(* IEC 61131-3 sources: 2026_Projet_YGO_ExcavatriceDragage/TOOLS/TEST_AUTO_CI/RESULTS/L_SIMULATION/tests (part 11) *)

TEST 'TC-T418-INT-010 Desactivation source pendant armement'
nx := 5000; ny := 5000; raw1 := 0; raw2 := 0; previousButton := FALSE; buttonEdges := 0;
bench.Enable := TRUE; bench.HwReal.Operator.JoyXRaw_ANA1 := 5000; bench.HwReal.Operator.JoyYRaw_ANA2 := 5000;
ADVANCE_TIME(10000000); bench(RawPosM1 := raw1, RawPosM2 := raw2);
bench.SimJoystickRight_Fwd_MAINT_Active := TRUE;
ADVANCE_TIME(10000000); bench(RawPosM1 := raw1, RawPosM2 := raw2);
ADVANCE_TIME(10000000); bench(RawPosM1 := raw1, RawPosM2 := raw2);
ADVANCE_TIME(10000000); bench(RawPosM1 := raw1, RawPosM2 := raw2);
ADVANCE_TIME(10000000); bench(RawPosM1 := raw1, RawPosM2 := raw2);
ADVANCE_TIME(10000000); bench(RawPosM1 := raw1, RawPosM2 := raw2);
ASSERT_TRUE(bench.Operator.JoyBtnRaw, 'Armement en cours');
bench.OperatorSourceActive := FALSE;
ADVANCE_TIME(10000000); bench(RawPosM1 := raw1, RawPosM2 := raw2);
ADVANCE_TIME(10000000); bench(RawPosM1 := raw1, RawPosM2 := raw2);
ADVANCE_TIME(10000000); bench(RawPosM1 := raw1, RawPosM2 := raw2);
ADVANCE_TIME(10000000); bench(RawPosM1 := raw1, RawPosM2 := raw2);
ADVANCE_TIME(10000000); bench(RawPosM1 := raw1, RawPosM2 := raw2);
ADVANCE_TIME(10000000); bench(RawPosM1 := raw1, RawPosM2 := raw2);
ADVANCE_TIME(10000000); bench(RawPosM1 := raw1, RawPosM2 := raw2);
ADVANCE_TIME(10000000); bench(RawPosM1 := raw1, RawPosM2 := raw2);
ADVANCE_TIME(10000000); bench(RawPosM1 := raw1, RawPosM2 := raw2);
ADVANCE_TIME(10000000); bench(RawPosM1 := raw1, RawPosM2 := raw2);
ASSERT_FALSE(bench.Operator.JoyBtnRaw, 'Source reelle sans bouton'); ASSERT_EQ(bench.Operator.JoyXRaw_ANA1, 5000, 'Neutre reel');
bench.OperatorSourceActive := TRUE;
ADVANCE_TIME(10000000); bench(RawPosM1 := raw1, RawPosM2 := raw2);
ADVANCE_TIME(10000000); bench(RawPosM1 := raw1, RawPosM2 := raw2);
ADVANCE_TIME(10000000); bench(RawPosM1 := raw1, RawPosM2 := raw2);
ADVANCE_TIME(10000000); bench(RawPosM1 := raw1, RawPosM2 := raw2);
ADVANCE_TIME(10000000); bench(RawPosM1 := raw1, RawPosM2 := raw2);
ADVANCE_TIME(10000000); bench(RawPosM1 := raw1, RawPosM2 := raw2);
ADVANCE_TIME(10000000); bench(RawPosM1 := raw1, RawPosM2 := raw2);
ADVANCE_TIME(10000000); bench(RawPosM1 := raw1, RawPosM2 := raw2);
ADVANCE_TIME(10000000); bench(RawPosM1 := raw1, RawPosM2 := raw2);
ADVANCE_TIME(10000000); bench(RawPosM1 := raw1, RawPosM2 := raw2);
ADVANCE_TIME(10000000); bench(RawPosM1 := raw1, RawPosM2 := raw2);
ADVANCE_TIME(10000000); bench(RawPosM1 := raw1, RawPosM2 := raw2);
ADVANCE_TIME(10000000); bench(RawPosM1 := raw1, RawPosM2 := raw2);
ADVANCE_TIME(10000000); bench(RawPosM1 := raw1, RawPosM2 := raw2);
ADVANCE_TIME(10000000); bench(RawPosM1 := raw1, RawPosM2 := raw2);
ADVANCE_TIME(10000000); bench(RawPosM1 := raw1, RawPosM2 := raw2);
ADVANCE_TIME(10000000); bench(RawPosM1 := raw1, RawPosM2 := raw2);
ADVANCE_TIME(10000000); bench(RawPosM1 := raw1, RawPosM2 := raw2);
ADVANCE_TIME(10000000); bench(RawPosM1 := raw1, RawPosM2 := raw2);
ADVANCE_TIME(10000000); bench(RawPosM1 := raw1, RawPosM2 := raw2);
ADVANCE_TIME(10000000); bench(RawPosM1 := raw1, RawPosM2 := raw2);
ADVANCE_TIME(10000000); bench(RawPosM1 := raw1, RawPosM2 := raw2);
ADVANCE_TIME(10000000); bench(RawPosM1 := raw1, RawPosM2 := raw2);
ADVANCE_TIME(10000000); bench(RawPosM1 := raw1, RawPosM2 := raw2);
ADVANCE_TIME(10000000); bench(RawPosM1 := raw1, RawPosM2 := raw2);
ADVANCE_TIME(10000000); bench(RawPosM1 := raw1, RawPosM2 := raw2);
ADVANCE_TIME(10000000); bench(RawPosM1 := raw1, RawPosM2 := raw2);
ADVANCE_TIME(10000000); bench(RawPosM1 := raw1, RawPosM2 := raw2);
ADVANCE_TIME(10000000); bench(RawPosM1 := raw1, RawPosM2 := raw2);
ADVANCE_TIME(10000000); bench(RawPosM1 := raw1, RawPosM2 := raw2);
ADVANCE_TIME(10000000); bench(RawPosM1 := raw1, RawPosM2 := raw2);
ADVANCE_TIME(10000000); bench(RawPosM1 := raw1, RawPosM2 := raw2);
ADVANCE_TIME(10000000); bench(RawPosM1 := raw1, RawPosM2 := raw2);
ADVANCE_TIME(10000000); bench(RawPosM1 := raw1, RawPosM2 := raw2);
ADVANCE_TIME(10000000); bench(RawPosM1 := raw1, RawPosM2 := raw2);
ADVANCE_TIME(10000000); bench(RawPosM1 := raw1, RawPosM2 := raw2);
ADVANCE_TIME(10000000); bench(RawPosM1 := raw1, RawPosM2 := raw2);
ADVANCE_TIME(10000000); bench(RawPosM1 := raw1, RawPosM2 := raw2);
ADVANCE_TIME(10000000); bench(RawPosM1 := raw1, RawPosM2 := raw2);
ADVANCE_TIME(10000000); bench(RawPosM1 := raw1, RawPosM2 := raw2);
ADVANCE_TIME(10000000); bench(RawPosM1 := raw1, RawPosM2 := raw2);
ADVANCE_TIME(10000000); bench(RawPosM1 := raw1, RawPosM2 := raw2);
ADVANCE_TIME(10000000); bench(RawPosM1 := raw1, RawPosM2 := raw2);
ADVANCE_TIME(10000000); bench(RawPosM1 := raw1, RawPosM2 := raw2);
ADVANCE_TIME(10000000); bench(RawPosM1 := raw1, RawPosM2 := raw2);
ADVANCE_TIME(10000000); bench(RawPosM1 := raw1, RawPosM2 := raw2);
ADVANCE_TIME(10000000); bench(RawPosM1 := raw1, RawPosM2 := raw2);
ADVANCE_TIME(10000000); bench(RawPosM1 := raw1, RawPosM2 := raw2);
ADVANCE_TIME(10000000); bench(RawPosM1 := raw1, RawPosM2 := raw2);
ADVANCE_TIME(10000000); bench(RawPosM1 := raw1, RawPosM2 := raw2);
ADVANCE_TIME(10000000); bench(RawPosM1 := raw1, RawPosM2 := raw2);
ADVANCE_TIME(10000000); bench(RawPosM1 := raw1, RawPosM2 := raw2);
ADVANCE_TIME(10000000); bench(RawPosM1 := raw1, RawPosM2 := raw2);
ADVANCE_TIME(10000000); bench(RawPosM1 := raw1, RawPosM2 := raw2);
ADVANCE_TIME(10000000); bench(RawPosM1 := raw1, RawPosM2 := raw2);
ADVANCE_TIME(10000000); bench(RawPosM1 := raw1, RawPosM2 := raw2);
ADVANCE_TIME(10000000); bench(RawPosM1 := raw1, RawPosM2 := raw2);
ADVANCE_TIME(10000000); bench(RawPosM1 := raw1, RawPosM2 := raw2);
ADVANCE_TIME(10000000); bench(RawPosM1 := raw1, RawPosM2 := raw2);
ADVANCE_TIME(10000000); bench(RawPosM1 := raw1, RawPosM2 := raw2);
ASSERT_FALSE(bench.Operator.JoyBtnRaw, 'Aucun rearmement apres retour de source'); ASSERT_EQ(bench.Operator.JoyXRaw_ANA1, 5000, 'IHM tenue ignoree');
bench.SimJoystickRight_Fwd_MAINT_Active := FALSE;
ADVANCE_TIME(10000000); bench(RawPosM1 := raw1, RawPosM2 := raw2);
bench.SimJoystickRight_Fwd_MAINT_Active := TRUE;
ADVANCE_TIME(10000000); bench(RawPosM1 := raw1, RawPosM2 := raw2);
ASSERT_TRUE(bench.Operator.JoyBtnRaw, 'Nouvel appui apres relachement disponible');
END_TEST

TEST 'TC-T418-INT-011 Desactivation source pendant retour'
nx := 5000; ny := 5000; raw1 := 0; raw2 := 0; previousButton := FALSE; buttonEdges := 0;
bench.Enable := TRUE; bench.HwReal.Operator.JoyXRaw_ANA1 := 5000; bench.HwReal.Operator.JoyYRaw_ANA2 := 5000;
ADVANCE_TIME(10000000); bench(RawPosM1 := raw1, RawPosM2 := raw2);
bench.SimJoystickRight_Fwd_MAINT_Active := TRUE;
ADVANCE_TIME(10000000); bench(RawPosM1 := raw1, RawPosM2 := raw2);
ADVANCE_TIME(10000000); bench(RawPosM1 := raw1, RawPosM2 := raw2);
ADVANCE_TIME(10000000); bench(RawPosM1 := raw1, RawPosM2 := raw2);
ADVANCE_TIME(10000000); bench(RawPosM1 := raw1, RawPosM2 := raw2);
ADVANCE_TIME(10000000); bench(RawPosM1 := raw1, RawPosM2 := raw2);
ADVANCE_TIME(10000000); bench(RawPosM1 := raw1, RawPosM2 := raw2);
ADVANCE_TIME(10000000); bench(RawPosM1 := raw1, RawPosM2 := raw2);
ADVANCE_TIME(10000000); bench(RawPosM1 := raw1, RawPosM2 := raw2);
ADVANCE_TIME(10000000); bench(RawPosM1 := raw1, RawPosM2 := raw2);
ADVANCE_TIME(10000000); bench(RawPosM1 := raw1, RawPosM2 := raw2);
ADVANCE_TIME(10000000); bench(RawPosM1 := raw1, RawPosM2 := raw2);
ADVANCE_TIME(10000000); bench(RawPosM1 := raw1, RawPosM2 := raw2);
ADVANCE_TIME(10000000); bench(RawPosM1 := raw1, RawPosM2 := raw2);
ADVANCE_TIME(10000000); bench(RawPosM1 := raw1, RawPosM2 := raw2);
ADVANCE_TIME(10000000); bench(RawPosM1 := raw1, RawPosM2 := raw2);
ADVANCE_TIME(10000000); bench(RawPosM1 := raw1, RawPosM2 := raw2);
ADVANCE_TIME(10000000); bench(RawPosM1 := raw1, RawPosM2 := raw2);
ADVANCE_TIME(10000000); bench(RawPosM1 := raw1, RawPosM2 := raw2);
ADVANCE_TIME(10000000); bench(RawPosM1 := raw1, RawPosM2 := raw2);
ADVANCE_TIME(10000000); bench(RawPosM1 := raw1, RawPosM2 := raw2);
ADVANCE_TIME(10000000); bench(RawPosM1 := raw1, RawPosM2 := raw2);
ADVANCE_TIME(10000000); bench(RawPosM1 := raw1, RawPosM2 := raw2);
ADVANCE_TIME(10000000); bench(RawPosM1 := raw1, RawPosM2 := raw2);
ADVANCE_TIME(10000000); bench(RawPosM1 := raw1, RawPosM2 := raw2);
ADVANCE_TIME(10000000); bench(RawPosM1 := raw1, RawPosM2 := raw2);
ADVANCE_TIME(10000000); bench(RawPosM1 := raw1, RawPosM2 := raw2);
ADVANCE_TIME(10000000); bench(RawPosM1 := raw1, RawPosM2 := raw2);
ADVANCE_TIME(10000000); bench(RawPosM1 := raw1, RawPosM2 := raw2);
ADVANCE_TIME(10000000); bench(RawPosM1 := raw1, RawPosM2 := raw2);
ADVANCE_TIME(10000000); bench(RawPosM1 := raw1, RawPosM2 := raw2);
ADVANCE_TIME(10000000); bench(RawPosM1 := raw1, RawPosM2 := raw2);
ADVANCE_TIME(10000000); bench(RawPosM1 := raw1, RawPosM2 := raw2);
ADVANCE_TIME(10000000); bench(RawPosM1 := raw1, RawPosM2 := raw2);
ADVANCE_TIME(10000000); bench(RawPosM1 := raw1, RawPosM2 := raw2);
ADVANCE_TIME(10000000); bench(RawPosM1 := raw1, RawPosM2 := raw2);
ADVANCE_TIME(10000000); bench(RawPosM1 := raw1, RawPosM2 := raw2);
ADVANCE_TIME(10000000); bench(RawPosM1 := raw1, RawPosM2 := raw2);
ADVANCE_TIME(10000000); bench(RawPosM1 := raw1, RawPosM2 := raw2);
ADVANCE_TIME(10000000); bench(RawPosM1 := raw1, RawPosM2 := raw2);
ADVANCE_TIME(10000000); bench(RawPosM1 := raw1, RawPosM2 := raw2);
ADVANCE_TIME(10000000); bench(RawPosM1 := raw1, RawPosM2 := raw2);
ADVANCE_TIME(10000000); bench(RawPosM1 := raw1, RawPosM2 := raw2);
ADVANCE_TIME(10000000); bench(RawPosM1 := raw1, RawPosM2 := raw2);
ADVANCE_TIME(10000000); bench(RawPosM1 := raw1, RawPosM2 := raw2);
ADVANCE_TIME(10000000); bench(RawPosM1 := raw1, RawPosM2 := raw2);
ADVANCE_TIME(10000000); bench(RawPosM1 := raw1, RawPosM2 := raw2);
ADVANCE_TIME(10000000); bench(RawPosM1 := raw1, RawPosM2 := raw2);
ADVANCE_TIME(10000000); bench(RawPosM1 := raw1, RawPosM2 := raw2);
ADVANCE_TIME(10000000); bench(RawPosM1 := raw1, RawPosM2 := raw2);
ADVANCE_TIME(10000000); bench(RawPosM1 := raw1, RawPosM2 := raw2);
ADVANCE_TIME(10000000); bench(RawPosM1 := raw1, RawPosM2 := raw2);
ADVANCE_TIME(10000000); bench(RawPosM1 := raw1, RawPosM2 := raw2);
ADVANCE_TIME(10000000); bench(RawPosM1 := raw1, RawPosM2 := raw2);
ADVANCE_TIME(10000000); bench(RawPosM1 := raw1, RawPosM2 := raw2);
ADVANCE_TIME(10000000); bench(RawPosM1 := raw1, RawPosM2 := raw2);
ADVANCE_TIME(10000000); bench(RawPosM1 := raw1, RawPosM2 := raw2);
ADVANCE_TIME(10000000); bench(RawPosM1 := raw1, RawPosM2 := raw2);
ADVANCE_TIME(10000000); bench(RawPosM1 := raw1, RawPosM2 := raw2);
ADVANCE_TIME(10000000); bench(RawPosM1 := raw1, RawPosM2 := raw2);
ADVANCE_TIME(10000000); bench(RawPosM1 := raw1, RawPosM2 := raw2);
ADVANCE_TIME(10000000); bench(RawPosM1 := raw1, RawPosM2 := raw2);
ADVANCE_TIME(10000000); bench(RawPosM1 := raw1, RawPosM2 := raw2);
ADVANCE_TIME(10000000); bench(RawPosM1 := raw1, RawPosM2 := raw2);
ADVANCE_TIME(10000000); bench(RawPosM1 := raw1, RawPosM2 := raw2);
ADVANCE_TIME(10000000); bench(RawPosM1 := raw1, RawPosM2 := raw2);
bench.SimJoystickRight_Fwd_MAINT_Active := FALSE;
ADVANCE_TIME(10000000); bench(RawPosM1 := raw1, RawPosM2 := raw2);
bench.OperatorSourceActive := FALSE;
ADVANCE_TIME(10000000); bench(RawPosM1 := raw1, RawPosM2 := raw2);
bench.SimJoystickLeft_Rev_TREMIE_Active := TRUE; bench.OperatorSourceActive := TRUE;
ADVANCE_TIME(10000000); bench(RawPosM1 := raw1, RawPosM2 := raw2);
ADVANCE_TIME(10000000); bench(RawPosM1 := raw1, RawPosM2 := raw2);
ADVANCE_TIME(10000000); bench(RawPosM1 := raw1, RawPosM2 := raw2);
ADVANCE_TIME(10000000); bench(RawPosM1 := raw1, RawPosM2 := raw2);
ADVANCE_TIME(10000000); bench(RawPosM1 := raw1, RawPosM2 := raw2);
ADVANCE_TIME(10000000); bench(RawPosM1 := raw1, RawPosM2 := raw2);
ADVANCE_TIME(10000000); bench(RawPosM1 := raw1, RawPosM2 := raw2);
ADVANCE_TIME(10000000); bench(RawPosM1 := raw1, RawPosM2 := raw2);
ADVANCE_TIME(10000000); bench(RawPosM1 := raw1, RawPosM2 := raw2);
ADVANCE_TIME(10000000); bench(RawPosM1 := raw1, RawPosM2 := raw2);
ADVANCE_TIME(10000000); bench(RawPosM1 := raw1, RawPosM2 := raw2);
ADVANCE_TIME(10000000); bench(RawPosM1 := raw1, RawPosM2 := raw2);
ADVANCE_TIME(10000000); bench(RawPosM1 := raw1, RawPosM2 := raw2);
ADVANCE_TIME(10000000); bench(RawPosM1 := raw1, RawPosM2 := raw2);
ADVANCE_TIME(10000000); bench(RawPosM1 := raw1, RawPosM2 := raw2);
ADVANCE_TIME(10000000); bench(RawPosM1 := raw1, RawPosM2 := raw2);
ADVANCE_TIME(10000000); bench(RawPosM1 := raw1, RawPosM2 := raw2);
ADVANCE_TIME(10000000); bench(RawPosM1 := raw1, RawPosM2 := raw2);
ADVANCE_TIME(10000000); bench(RawPosM1 := raw1, RawPosM2 := raw2);
ADVANCE_TIME(10000000); bench(RawPosM1 := raw1, RawPosM2 := raw2);
ADVANCE_TIME(10000000); bench(RawPosM1 := raw1, RawPosM2 := raw2);
ADVANCE_TIME(10000000); bench(RawPosM1 := raw1, RawPosM2 := raw2);
ADVANCE_TIME(10000000); bench(RawPosM1 := raw1, RawPosM2 := raw2);
ADVANCE_TIME(10000000); bench(RawPosM1 := raw1, RawPosM2 := raw2);
ADVANCE_TIME(10000000); bench(RawPosM1 := raw1, RawPosM2 := raw2);
ADVANCE_TIME(10000000); bench(RawPosM1 := raw1, RawPosM2 := raw2);
ADVANCE_TIME(10000000); bench(RawPosM1 := raw1, RawPosM2 := raw2);
ADVANCE_TIME(10000000); bench(RawPosM1 := raw1, RawPosM2 := raw2);
ADVANCE_TIME(10000000); bench(RawPosM1 := raw1, RawPosM2 := raw2);
ADVANCE_TIME(10000000); bench(RawPosM1 := raw1, RawPosM2 := raw2);
ADVANCE_TIME(10000000); bench(RawPosM1 := raw1, RawPosM2 := raw2);
ADVANCE_TIME(10000000); bench(RawPosM1 := raw1, RawPosM2 := raw2);
ADVANCE_TIME(10000000); bench(RawPosM1 := raw1, RawPosM2 := raw2);
ADVANCE_TIME(10000000); bench(RawPosM1 := raw1, RawPosM2 := raw2);
ADVANCE_TIME(10000000); bench(RawPosM1 := raw1, RawPosM2 := raw2);
ADVANCE_TIME(10000000); bench(RawPosM1 := raw1, RawPosM2 := raw2);
ADVANCE_TIME(10000000); bench(RawPosM1 := raw1, RawPosM2 := raw2);
ADVANCE_TIME(10000000); bench(RawPosM1 := raw1, RawPosM2 := raw2);
ADVANCE_TIME(10000000); bench(RawPosM1 := raw1, RawPosM2 := raw2);
ADVANCE_TIME(10000000); bench(RawPosM1 := raw1, RawPosM2 := raw2);
ADVANCE_TIME(10000000); bench(RawPosM1 := raw1, RawPosM2 := raw2);
ADVANCE_TIME(10000000); bench(RawPosM1 := raw1, RawPosM2 := raw2);
ADVANCE_TIME(10000000); bench(RawPosM1 := raw1, RawPosM2 := raw2);
ADVANCE_TIME(10000000); bench(RawPosM1 := raw1, RawPosM2 := raw2);
ADVANCE_TIME(10000000); bench(RawPosM1 := raw1, RawPosM2 := raw2);
ADVANCE_TIME(10000000); bench(RawPosM1 := raw1, RawPosM2 := raw2);
ADVANCE_TIME(10000000); bench(RawPosM1 := raw1, RawPosM2 := raw2);
ADVANCE_TIME(10000000); bench(RawPosM1 := raw1, RawPosM2 := raw2);
ADVANCE_TIME(10000000); bench(RawPosM1 := raw1, RawPosM2 := raw2);
ADVANCE_TIME(10000000); bench(RawPosM1 := raw1, RawPosM2 := raw2);
ADVANCE_TIME(10000000); bench(RawPosM1 := raw1, RawPosM2 := raw2);
ADVANCE_TIME(10000000); bench(RawPosM1 := raw1, RawPosM2 := raw2);
ADVANCE_TIME(10000000); bench(RawPosM1 := raw1, RawPosM2 := raw2);
ADVANCE_TIME(10000000); bench(RawPosM1 := raw1, RawPosM2 := raw2);
ADVANCE_TIME(10000000); bench(RawPosM1 := raw1, RawPosM2 := raw2);
ADVANCE_TIME(10000000); bench(RawPosM1 := raw1, RawPosM2 := raw2);
ADVANCE_TIME(10000000); bench(RawPosM1 := raw1, RawPosM2 := raw2);
ADVANCE_TIME(10000000); bench(RawPosM1 := raw1, RawPosM2 := raw2);
ADVANCE_TIME(10000000); bench(RawPosM1 := raw1, RawPosM2 := raw2);
ADVANCE_TIME(10000000); bench(RawPosM1 := raw1, RawPosM2 := raw2);
ASSERT_EQ(bench.Operator.JoyXRaw_ANA1, 5000, 'Retour interrompu ne charge aucun nouveau geste'); ASSERT_FALSE(bench.Operator.JoyBtnRaw, 'Aucun appui differe');
END_TEST

TEST 'TC-T418-INT-012 Source reelle restitue image sans stimuli manuels'
nx := 5000; ny := 5000; raw1 := 0; raw2 := 0; previousButton := FALSE; buttonEdges := 0;
bench.Enable := TRUE; bench.HwReal.Operator.JoyXRaw_ANA1 := 5000; bench.HwReal.Operator.JoyYRaw_ANA2 := 5000;
bench.OperatorSourceActive := FALSE; bench.SimJoystickRawX := 9999; bench.SimJoystickRawY := 1; bench.SimJoystickRawButton := TRUE;
bench.HwReal.Operator.JoyXRaw_ANA1 := 4321; bench.HwReal.Operator.JoyYRaw_ANA2 := 6789; bench.HwReal.Operator.JoyBtnRaw := FALSE; bench.HwReal.Operator.CanBusState := 0;
ADVANCE_TIME(10000000); bench(RawPosM1 := raw1, RawPosM2 := raw2);
ASSERT_EQ(bench.Operator.JoyXRaw_ANA1, 4321, 'X reel exact'); ASSERT_EQ(bench.Operator.JoyYRaw_ANA2, 6789, 'Y reel exact'); ASSERT_FALSE(bench.Operator.JoyBtnRaw, 'Bouton reel exact'); ASSERT_EQ(bench.Operator.CanBusState, 0, 'Diagnostic reel non remplace par RUNNING');
END_TEST

(* ---- test_sim_translation_loop.st ---- *)
(* T417 - rejeu en boucle fermee : FB_Translation REEL (non modifie) + decodeur + FB_Sim_Translation.
   Voir MOCKS/FB_TestLoopTranslation.st (cablage PRG_05 reproduit ; FB_TranslationOutputInterlock et
   FB_Safety_Translation NON reproduits). Un scan = 20 ms simules. Tests de CARACTERISATION : bandes larges,
   gain 0,02 m/(Hz.s) provisoire (T301) ; ce ne sont pas des mesures terrain. *)

TEST 'TC-T417-LOOP-A Rejeu P1 a 20 Hz, demande TENUE apres arrivee : le plafond d approche maintient 20 Hz vers le variateur'
VAR
    loop : FB_TestLoopTranslation;
END_VAR
    loop.HoldRequest := TRUE;
    ADVANCE_TIME(20000000); loop();
    ADVANCE_TIME(20000000); loop();
    ADVANCE_TIME(20000000); loop();
    ADVANCE_TIME(20000000); loop();
    ADVANCE_TIME(20000000); loop();
    ADVANCE_TIME(20000000); loop();
    ADVANCE_TIME(20000000); loop();
    ADVANCE_TIME(20000000); loop();
    ADVANCE_TIME(20000000); loop();
    ADVANCE_TIME(20000000); loop();
    ADVANCE_TIME(20000000); loop();
    ADVANCE_TIME(20000000); loop();
    ADVANCE_TIME(20000000); loop();
    ADVANCE_TIME(20000000); loop();
    ADVANCE_TIME(20000000); loop();
    ADVANCE_TIME(20000000); loop();
    ADVANCE_TIME(20000000); loop();
    ADVANCE_TIME(20000000); loop();
    ADVANCE_TIME(20000000); loop();
    ADVANCE_TIME(20000000); loop();
    ADVANCE_TIME(20000000); loop();
    ADVANCE_TIME(20000000); loop();
    ADVANCE_TIME(20000000); loop();
    ADVANCE_TIME(20000000); loop();
    ADVANCE_TIME(20000000); loop();
    ADVANCE_TIME(20000000); loop();
    ADVANCE_TIME(20000000); loop();
    ADVANCE_TIME(20000000); loop();
    ADVANCE_TIME(20000000); loop();
    ADVANCE_TIME(20000000); loop();
    ADVANCE_TIME(20000000); loop();
    ADVANCE_TIME(20000000); loop();
    ADVANCE_TIME(20000000); loop();
    ADVANCE_TIME(20000000); loop();
    ADVANCE_TIME(20000000); loop();
    ADVANCE_TIME(20000000); loop();
    ADVANCE_TIME(20000000); loop();
    ADVANCE_TIME(20000000); loop();
    ADVANCE_TIME(20000000); loop();
    ADVANCE_TIME(20000000); loop();
    ADVANCE_TIME(20000000); loop();
    ADVANCE_TIME(20000000); loop();
    ADVANCE_TIME(20000000); loop();
    ADVANCE_TIME(20000000); loop();
    ADVANCE_TIME(20000000); loop();
    ADVANCE_TIME(20000000); loop();
    ADVANCE_TIME(20000000); loop();
    ADVANCE_TIME(20000000); loop();
    ADVANCE_TIME(20000000); loop();
    ADVANCE_TIME(20000000); loop();
    ADVANCE_TIME(20000000); loop();
    ADVANCE_TIME(20000000); loop();
    ADVANCE_TIME(20000000); loop();
    ADVANCE_TIME(20000000); loop();
    ADVANCE_TIME(20000000); loop();
    ADVANCE_TIME(20000000); loop();
    ADVANCE_TIME(20000000); loop();
    ADVANCE_TIME(20000000); loop();
    ADVANCE_TIME(20000000); loop();
    ADVANCE_TIME(20000000); loop();
    ADVANCE_TIME(20000000); loop();
    ADVANCE_TIME(20000000); loop();
    ADVANCE_TIME(20000000); loop();
    ADVANCE_TIME(20000000); loop();
    ADVANCE_TIME(20000000); loop();
    ADVANCE_TIME(20000000); loop();
    ADVANCE_TIME(20000000); loop();
    ADVANCE_TIME(20000000); loop();
    ADVANCE_TIME(20000000); loop();
    ADVANCE_TIME(20000000); loop();
    ADVANCE_TIME(20000000); loop();
    ADVANCE_TIME(20000000); loop();
    ADVANCE_TIME(20000000); loop();
    ADVANCE_TIME(20000000); loop();
    ADVANCE_TIME(20000000); loop();
    ADVANCE_TIME(20000000); loop();
    ADVANCE_TIME(20000000); loop();
    ADVANCE_TIME(20000000); loop();
    ADVANCE_TIME(20000000); loop();
    ADVANCE_TIME(20000000); loop();
    ADVANCE_TIME(20000000); loop();
    ADVANCE_TIME(20000000); loop();
    ADVANCE_TIME(20000000); loop();
    ADVANCE_TIME(20000000); loop();
    ADVANCE_TIME(20000000); loop();
    ADVANCE_TIME(20000000); loop();
    ADVANCE_TIME(20000000); loop();
    ADVANCE_TIME(20000000); loop();
    ADVANCE_TIME(20000000); loop();
    ADVANCE_TIME(20000000); loop();
    ADVANCE_TIME(20000000); loop();
    ADVANCE_TIME(20000000); loop();
    ADVANCE_TIME(20000000); loop();
    ADVANCE_TIME(20000000); loop();
    ADVANCE_TIME(20000000); loop();
    ADVANCE_TIME(20000000); loop();
    ADVANCE_TIME(20000000); loop();
    ADVANCE_TIME(20000000); loop();
    ADVANCE_TIME(20000000); loop();
    ADVANCE_TIME(20000000); loop();
    ADVANCE_TIME(20000000); loop();
    ADVANCE_TIME(20000000); loop();
    ADVANCE_TIME(20000000); loop();
    ADVANCE_TIME(20000000); loop();
    ADVANCE_TIME(20000000); loop();
    ADVANCE_TIME(20000000); loop();
    ADVANCE_TIME(20000000); loop();
    ADVANCE_TIME(20000000); loop();
    ADVANCE_TIME(20000000); loop();
    ADVANCE_TIME(20000000); loop();
    ADVANCE_TIME(20000000); loop();
    ADVANCE_TIME(20000000); loop();
    ADVANCE_TIME(20000000); loop();
    ADVANCE_TIME(20000000); loop();
    ADVANCE_TIME(20000000); loop();
    ADVANCE_TIME(20000000); loop();
    ADVANCE_TIME(20000000); loop();
    ADVANCE_TIME(20000000); loop();
    ADVANCE_TIME(20000000); loop();
    ADVANCE_TIME(20000000); loop();
    ADVANCE_TIME(20000000); loop();
    ADVANCE_TIME(20000000); loop();
    ADVANCE_TIME(20000000); loop();
    ADVANCE_TIME(20000000); loop();
    ADVANCE_TIME(20000000); loop();
    ADVANCE_TIME(20000000); loop();
    ADVANCE_TIME(20000000); loop();
    ADVANCE_TIME(20000000); loop();
    ADVANCE_TIME(20000000); loop();
    ADVANCE_TIME(20000000); loop();
    ADVANCE_TIME(20000000); loop();
    ADVANCE_TIME(20000000); loop();
    ADVANCE_TIME(20000000); loop();
    ADVANCE_TIME(20000000); loop();
    ADVANCE_TIME(20000000); loop();
    ADVANCE_TIME(20000000); loop();
    ADVANCE_TIME(20000000); loop();
    ADVANCE_TIME(20000000); loop();
    ADVANCE_TIME(20000000); loop();
    ADVANCE_TIME(20000000); loop();
    ADVANCE_TIME(20000000); loop();
    ADVANCE_TIME(20000000); loop();
    ADVANCE_TIME(20000000); loop();
    ADVANCE_TIME(20000000); loop();
    ADVANCE_TIME(20000000); loop();
    ADVANCE_TIME(20000000); loop();
    ADVANCE_TIME(20000000); loop();
    ADVANCE_TIME(20000000); loop();
    ADVANCE_TIME(20000000); loop();
    ADVANCE_TIME(20000000); loop();
    ADVANCE_TIME(20000000); loop();
    ADVANCE_TIME(20000000); loop();
    ADVANCE_TIME(20000000); loop();
    ADVANCE_TIME(20000000); loop();
    ADVANCE_TIME(20000000); loop();
    ADVANCE_TIME(20000000); loop();
    ADVANCE_TIME(20000000); loop();
    ADVANCE_TIME(20000000); loop();
    ADVANCE_TIME(20000000); loop();
    ADVANCE_TIME(20000000); loop();
    ADVANCE_TIME(20000000); loop();
    ADVANCE_TIME(20000000); loop();
    ADVANCE_TIME(20000000); loop();
    ADVANCE_TIME(20000000); loop();
    ADVANCE_TIME(20000000); loop();
    ADVANCE_TIME(20000000); loop();
    ADVANCE_TIME(20000000); loop();
    ADVANCE_TIME(20000000); loop();
    ADVANCE_TIME(20000000); loop();
    ADVANCE_TIME(20000000); loop();
    ADVANCE_TIME(20000000); loop();
    ADVANCE_TIME(20000000); loop();
    ADVANCE_TIME(20000000); loop();
    ADVANCE_TIME(20000000); loop();
    ADVANCE_TIME(20000000); loop();
    ADVANCE_TIME(20000000); loop();
    ADVANCE_TIME(20000000); loop();
    ADVANCE_TIME(20000000); loop();
    ADVANCE_TIME(20000000); loop();
    ADVANCE_TIME(20000000); loop();
    ADVANCE_TIME(20000000); loop();
    ADVANCE_TIME(20000000); loop();
    ADVANCE_TIME(20000000); loop();
    ADVANCE_TIME(20000000); loop();
    ADVANCE_TIME(20000000); loop();
    ADVANCE_TIME(20000000); loop();
    ADVANCE_TIME(20000000); loop();
    ADVANCE_TIME(20000000); loop();
    ADVANCE_TIME(20000000); loop();
    ADVANCE_TIME(20000000); loop();
    ADVANCE_TIME(20000000); loop();
    ADVANCE_TIME(20000000); loop();
    ADVANCE_TIME(20000000); loop();
    ADVANCE_TIME(20000000); loop();
    ADVANCE_TIME(20000000); loop();
    ADVANCE_TIME(20000000); loop();
    ADVANCE_TIME(20000000); loop();
    ADVANCE_TIME(20000000); loop();
    ADVANCE_TIME(20000000); loop();
    ADVANCE_TIME(20000000); loop();
    ADVANCE_TIME(20000000); loop();
    ADVANCE_TIME(20000000); loop();
    ADVANCE_TIME(20000000); loop();
    ADVANCE_TIME(20000000); loop();
    ADVANCE_TIME(20000000); loop();
    ADVANCE_TIME(20000000); loop();
    ADVANCE_TIME(20000000); loop();
    ADVANCE_TIME(20000000); loop();
    ADVANCE_TIME(20000000); loop();
    ADVANCE_TIME(20000000); loop();
    ADVANCE_TIME(20000000); loop();
    ADVANCE_TIME(20000000); loop();
    ADVANCE_TIME(20000000); loop();
    ADVANCE_TIME(20000000); loop();
    ADVANCE_TIME(20000000); loop();
    ADVANCE_TIME(20000000); loop();
    ADVANCE_TIME(20000000); loop();
    ADVANCE_TIME(20000000); loop();
    ADVANCE_TIME(20000000); loop();
    ADVANCE_TIME(20000000); loop();
    ADVANCE_TIME(20000000); loop();
    ADVANCE_TIME(20000000); loop();
    ADVANCE_TIME(20000000); loop();
    ADVANCE_TIME(20000000); loop();
    ADVANCE_TIME(20000000); loop();
    ADVANCE_TIME(20000000); loop();
    ADVANCE_TIME(20000000); loop();
    ADVANCE_TIME(20000000); loop();
    ADVANCE_TIME(20000000); loop();
    ADVANCE_TIME(20000000); loop();
    ADVANCE_TIME(20000000); loop();
    ADVANCE_TIME(20000000); loop();
    ADVANCE_TIME(20000000); loop();
    ADVANCE_TIME(20000000); loop();
    ADVANCE_TIME(20000000); loop();
    ADVANCE_TIME(20000000); loop();
    ADVANCE_TIME(20000000); loop();
    ADVANCE_TIME(20000000); loop();
    ADVANCE_TIME(20000000); loop();
    ADVANCE_TIME(20000000); loop();
    ADVANCE_TIME(20000000); loop();
    ADVANCE_TIME(20000000); loop();
    ADVANCE_TIME(20000000); loop();
    ADVANCE_TIME(20000000); loop();
    ADVANCE_TIME(20000000); loop();
    ADVANCE_TIME(20000000); loop();
    ADVANCE_TIME(20000000); loop();
    ADVANCE_TIME(20000000); loop();
    ADVANCE_TIME(20000000); loop();
    ADVANCE_TIME(20000000); loop();
    ADVANCE_TIME(20000000); loop();
    ADVANCE_TIME(20000000); loop();
    ADVANCE_TIME(20000000); loop();
    ADVANCE_TIME(20000000); loop();
    ADVANCE_TIME(20000000); loop();
    ADVANCE_TIME(20000000); loop();
    ADVANCE_TIME(20000000); loop();
    ADVANCE_TIME(20000000); loop();
    ADVANCE_TIME(20000000); loop();
    ADVANCE_TIME(20000000); loop();
    ADVANCE_TIME(20000000); loop();
    ADVANCE_TIME(20000000); loop();
    ADVANCE_TIME(20000000); loop();
    ADVANCE_TIME(20000000); loop();
    ADVANCE_TIME(20000000); loop();
    ADVANCE_TIME(20000000); loop();
    ADVANCE_TIME(20000000); loop();
    ADVANCE_TIME(20000000); loop();
    ADVANCE_TIME(20000000); loop();
    ADVANCE_TIME(20000000); loop();
    ADVANCE_TIME(20000000); loop();
    ADVANCE_TIME(20000000); loop();
    ADVANCE_TIME(20000000); loop();
    ADVANCE_TIME(20000000); loop();
    ADVANCE_TIME(20000000); loop();
    ADVANCE_TIME(20000000); loop();
    ADVANCE_TIME(20000000); loop();
    ADVANCE_TIME(20000000); loop();
    ADVANCE_TIME(20000000); loop();
    ADVANCE_TIME(20000000); loop();
    ADVANCE_TIME(20000000); loop();
    ADVANCE_TIME(20000000); loop();
    ADVANCE_TIME(20000000); loop();
    ADVANCE_TIME(20000000); loop();
    ADVANCE_TIME(20000000); loop();
    ADVANCE_TIME(20000000); loop();
    ADVANCE_TIME(20000000); loop();
    ADVANCE_TIME(20000000); loop();
    ADVANCE_TIME(20000000); loop();
    ADVANCE_TIME(20000000); loop();
    ADVANCE_TIME(20000000); loop();
    ADVANCE_TIME(20000000); loop();
    ADVANCE_TIME(20000000); loop();
    ADVANCE_TIME(20000000); loop();
    ADVANCE_TIME(20000000); loop();
    ADVANCE_TIME(20000000); loop();
    ADVANCE_TIME(20000000); loop();
    ADVANCE_TIME(20000000); loop();
    ADVANCE_TIME(20000000); loop();
    ADVANCE_TIME(20000000); loop();
    ADVANCE_TIME(20000000); loop();
    ADVANCE_TIME(20000000); loop();
    ADVANCE_TIME(20000000); loop();
    ADVANCE_TIME(20000000); loop();
    ADVANCE_TIME(20000000); loop();
    ADVANCE_TIME(20000000); loop();
    ADVANCE_TIME(20000000); loop();
    ADVANCE_TIME(20000000); loop();
    ADVANCE_TIME(20000000); loop();
    ADVANCE_TIME(20000000); loop();
    ADVANCE_TIME(20000000); loop();
    ADVANCE_TIME(20000000); loop();
    ADVANCE_TIME(20000000); loop();
    ADVANCE_TIME(20000000); loop();
    ADVANCE_TIME(20000000); loop();
    ADVANCE_TIME(20000000); loop();
    ADVANCE_TIME(20000000); loop();
    ADVANCE_TIME(20000000); loop();
    ADVANCE_TIME(20000000); loop();
    ADVANCE_TIME(20000000); loop();
    ADVANCE_TIME(20000000); loop();
    ADVANCE_TIME(20000000); loop();
    ADVANCE_TIME(20000000); loop();
    ADVANCE_TIME(20000000); loop();
    ADVANCE_TIME(20000000); loop();
    ADVANCE_TIME(20000000); loop();
    ADVANCE_TIME(20000000); loop();
    ADVANCE_TIME(20000000); loop();
    ADVANCE_TIME(20000000); loop();
    ADVANCE_TIME(20000000); loop();
    ADVANCE_TIME(20000000); loop();
    ADVANCE_TIME(20000000); loop();
    ADVANCE_TIME(20000000); loop();
    ADVANCE_TIME(20000000); loop();
    ADVANCE_TIME(20000000); loop();
    ADVANCE_TIME(20000000); loop();
    ADVANCE_TIME(20000000); loop();
    ADVANCE_TIME(20000000); loop();
    ADVANCE_TIME(20000000); loop();
    ADVANCE_TIME(20000000); loop();
    ADVANCE_TIME(20000000); loop();
    ADVANCE_TIME(20000000); loop();
    ADVANCE_TIME(20000000); loop();
    ADVANCE_TIME(20000000); loop();
    ADVANCE_TIME(20000000); loop();
    ADVANCE_TIME(20000000); loop();
    ADVANCE_TIME(20000000); loop();
    ADVANCE_TIME(20000000); loop();
    ADVANCE_TIME(20000000); loop();
    ADVANCE_TIME(20000000); loop();
    ADVANCE_TIME(20000000); loop();
    ADVANCE_TIME(20000000); loop();
    ADVANCE_TIME(20000000); loop();
    ADVANCE_TIME(20000000); loop();
    ADVANCE_TIME(20000000); loop();
    ADVANCE_TIME(20000000); loop();
    ADVANCE_TIME(20000000); loop();
    ADVANCE_TIME(20000000); loop();
    ADVANCE_TIME(20000000); loop();
    ADVANCE_TIME(20000000); loop();
    ADVANCE_TIME(20000000); loop();
    ADVANCE_TIME(20000000); loop();
    ADVANCE_TIME(20000000); loop();
    ADVANCE_TIME(20000000); loop();
    ADVANCE_TIME(20000000); loop();
    ADVANCE_TIME(20000000); loop();
    ADVANCE_TIME(20000000); loop();
    ADVANCE_TIME(20000000); loop();
    ADVANCE_TIME(20000000); loop();
    ADVANCE_TIME(20000000); loop();
    ADVANCE_TIME(20000000); loop();
    ADVANCE_TIME(20000000); loop();
    ADVANCE_TIME(20000000); loop();
    ADVANCE_TIME(20000000); loop();
    ADVANCE_TIME(20000000); loop();
    ADVANCE_TIME(20000000); loop();
    ADVANCE_TIME(20000000); loop();
    ADVANCE_TIME(20000000); loop();
    ADVANCE_TIME(20000000); loop();
    ADVANCE_TIME(20000000); loop();
    ADVANCE_TIME(20000000); loop();
    ADVANCE_TIME(20000000); loop();
    ADVANCE_TIME(20000000); loop();
    ADVANCE_TIME(20000000); loop();
    ADVANCE_TIME(20000000); loop();
    ADVANCE_TIME(20000000); loop();
    ADVANCE_TIME(20000000); loop();
    ADVANCE_TIME(20000000); loop();
    ADVANCE_TIME(20000000); loop();
    ADVANCE_TIME(20000000); loop();
    ADVANCE_TIME(20000000); loop();
    ADVANCE_TIME(20000000); loop();
    ADVANCE_TIME(20000000); loop();
    ADVANCE_TIME(20000000); loop();
    ADVANCE_TIME(20000000); loop();
    ADVANCE_TIME(20000000); loop();
    ADVANCE_TIME(20000000); loop();
    ADVANCE_TIME(20000000); loop();
    ADVANCE_TIME(20000000); loop();
    ADVANCE_TIME(20000000); loop();
    ADVANCE_TIME(20000000); loop();
    ADVANCE_TIME(20000000); loop();
    ADVANCE_TIME(20000000); loop();
    ADVANCE_TIME(20000000); loop();
    ADVANCE_TIME(20000000); loop();
    ADVANCE_TIME(20000000); loop();
    ADVANCE_TIME(20000000); loop();
    ADVANCE_TIME(20000000); loop();
    ADVANCE_TIME(20000000); loop();
    ADVANCE_TIME(20000000); loop();
    ADVANCE_TIME(20000000); loop();
    ADVANCE_TIME(20000000); loop();
    ADVANCE_TIME(20000000); loop();
    ADVANCE_TIME(20000000); loop();
    ADVANCE_TIME(20000000); loop();
    ADVANCE_TIME(20000000); loop();
    ADVANCE_TIME(20000000); loop();
    ADVANCE_TIME(20000000); loop();
    ADVANCE_TIME(20000000); loop();
    ADVANCE_TIME(20000000); loop();
    ADVANCE_TIME(20000000); loop();
    ADVANCE_TIME(20000000); loop();
    ADVANCE_TIME(20000000); loop();
    ADVANCE_TIME(20000000); loop();
    ADVANCE_TIME(20000000); loop();
    ADVANCE_TIME(20000000); loop();
    ADVANCE_TIME(20000000); loop();
    ADVANCE_TIME(20000000); loop();
    ADVANCE_TIME(20000000); loop();
    ADVANCE_TIME(20000000); loop();
    ADVANCE_TIME(20000000); loop();
    ADVANCE_TIME(20000000); loop();
    ADVANCE_TIME(20000000); loop();
    ADVANCE_TIME(20000000); loop();
    ADVANCE_TIME(20000000); loop();
    ADVANCE_TIME(20000000); loop();
    ADVANCE_TIME(20000000); loop();
    ADVANCE_TIME(20000000); loop();
    ADVANCE_TIME(20000000); loop();
    ADVANCE_TIME(20000000); loop();
    ADVANCE_TIME(20000000); loop();
    ADVANCE_TIME(20000000); loop();
    ADVANCE_TIME(20000000); loop();
    ADVANCE_TIME(20000000); loop();
    ADVANCE_TIME(20000000); loop();
    ADVANCE_TIME(20000000); loop();
    ADVANCE_TIME(20000000); loop();
    ADVANCE_TIME(20000000); loop();
    ADVANCE_TIME(20000000); loop();
    ADVANCE_TIME(20000000); loop();
    ADVANCE_TIME(20000000); loop();
    ADVANCE_TIME(20000000); loop();
    ADVANCE_TIME(20000000); loop();
    ADVANCE_TIME(20000000); loop();
    ADVANCE_TIME(20000000); loop();
    ADVANCE_TIME(20000000); loop();
    ADVANCE_TIME(20000000); loop();
    ADVANCE_TIME(20000000); loop();
    ADVANCE_TIME(20000000); loop();
    ADVANCE_TIME(20000000); loop();
    ADVANCE_TIME(20000000); loop();
    ADVANCE_TIME(20000000); loop();
    ADVANCE_TIME(20000000); loop();
    ADVANCE_TIME(20000000); loop();
    ADVANCE_TIME(20000000); loop();
    ADVANCE_TIME(20000000); loop();
    ADVANCE_TIME(20000000); loop();
    ADVANCE_TIME(20000000); loop();
    ADVANCE_TIME(20000000); loop();
    ADVANCE_TIME(20000000); loop();
    ADVANCE_TIME(20000000); loop();
    ADVANCE_TIME(20000000); loop();
    ADVANCE_TIME(20000000); loop();
    ADVANCE_TIME(20000000); loop();
    ADVANCE_TIME(20000000); loop();
    ADVANCE_TIME(20000000); loop();
    ADVANCE_TIME(20000000); loop();
    ADVANCE_TIME(20000000); loop();
    ADVANCE_TIME(20000000); loop();
    ADVANCE_TIME(20000000); loop();
    ADVANCE_TIME(20000000); loop();
    ADVANCE_TIME(20000000); loop();
    ADVANCE_TIME(20000000); loop();
    ADVANCE_TIME(20000000); loop();
    ADVANCE_TIME(20000000); loop();
    ADVANCE_TIME(20000000); loop();
    ADVANCE_TIME(20000000); loop();
    ADVANCE_TIME(20000000); loop();
    ADVANCE_TIME(20000000); loop();
    ADVANCE_TIME(20000000); loop();
    ADVANCE_TIME(20000000); loop();
    ADVANCE_TIME(20000000); loop();
    ADVANCE_TIME(20000000); loop();
    ADVANCE_TIME(20000000); loop();
    ADVANCE_TIME(20000000); loop();
    ADVANCE_TIME(20000000); loop();
    ADVANCE_TIME(20000000); loop();
    ADVANCE_TIME(20000000); loop();
    ADVANCE_TIME(20000000); loop();
    ADVANCE_TIME(20000000); loop();
    ADVANCE_TIME(20000000); loop();
    ADVANCE_TIME(20000000); loop();
    ADVANCE_TIME(20000000); loop();
    ADVANCE_TIME(20000000); loop();
    ADVANCE_TIME(20000000); loop();
    ADVANCE_TIME(20000000); loop();
    ADVANCE_TIME(20000000); loop();
    ADVANCE_TIME(20000000); loop();
    ADVANCE_TIME(20000000); loop();
    ADVANCE_TIME(20000000); loop();
    ADVANCE_TIME(20000000); loop();
    ADVANCE_TIME(20000000); loop();
    ADVANCE_TIME(20000000); loop();
    ADVANCE_TIME(20000000); loop();
    ADVANCE_TIME(20000000); loop();
    ADVANCE_TIME(20000000); loop();
    ADVANCE_TIME(20000000); loop();
    ADVANCE_TIME(20000000); loop();
    ADVANCE_TIME(20000000); loop();
    ADVANCE_TIME(20000000); loop();
    ADVANCE_TIME(20000000); loop();
    ADVANCE_TIME(20000000); loop();
    ADVANCE_TIME(20000000); loop();
    ADVANCE_TIME(20000000); loop();
    ADVANCE_TIME(20000000); loop();
    ADVANCE_TIME(20000000); loop();
    ADVANCE_TIME(20000000); loop();
    ADVANCE_TIME(20000000); loop();
    ADVANCE_TIME(20000000); loop();
    ADVANCE_TIME(20000000); loop();
    ADVANCE_TIME(20000000); loop();
    ADVANCE_TIME(20000000); loop();
    ADVANCE_TIME(20000000); loop();
    ADVANCE_TIME(20000000); loop();
    ADVANCE_TIME(20000000); loop();
    ADVANCE_TIME(20000000); loop();
    ADVANCE_TIME(20000000); loop();
    ADVANCE_TIME(20000000); loop();
    ADVANCE_TIME(20000000); loop();
    ADVANCE_TIME(20000000); loop();
    ADVANCE_TIME(20000000); loop();
    ADVANCE_TIME(20000000); loop();
    ADVANCE_TIME(20000000); loop();
    ADVANCE_TIME(20000000); loop();
    ADVANCE_TIME(20000000); loop();
    ADVANCE_TIME(20000000); loop();
    ADVANCE_TIME(20000000); loop();
    ADVANCE_TIME(20000000); loop();
    ADVANCE_TIME(20000000); loop();
    ADVANCE_TIME(20000000); loop();
    ADVANCE_TIME(20000000); loop();
    ADVANCE_TIME(20000000); loop();
    ADVANCE_TIME(20000000); loop();
    ADVANCE_TIME(20000000); loop();
    ADVANCE_TIME(20000000); loop();
    ADVANCE_TIME(20000000); loop();
    ADVANCE_TIME(20000000); loop();
    ADVANCE_TIME(20000000); loop();
    ADVANCE_TIME(20000000); loop();
    ADVANCE_TIME(20000000); loop();
    ADVANCE_TIME(20000000); loop();
    ADVANCE_TIME(20000000); loop();
    ADVANCE_TIME(20000000); loop();
    ADVANCE_TIME(20000000); loop();
    ADVANCE_TIME(20000000); loop();
    ADVANCE_TIME(20000000); loop();
    ADVANCE_TIME(20000000); loop();
    ADVANCE_TIME(20000000); loop();
    ADVANCE_TIME(20000000); loop();
    ADVANCE_TIME(20000000); loop();
    ADVANCE_TIME(20000000); loop();
    ADVANCE_TIME(20000000); loop();
    ADVANCE_TIME(20000000); loop();
    ADVANCE_TIME(20000000); loop();
    ADVANCE_TIME(20000000); loop();
    ADVANCE_TIME(20000000); loop();
    ADVANCE_TIME(20000000); loop();
    ADVANCE_TIME(20000000); loop();
    ADVANCE_TIME(20000000); loop();
    ADVANCE_TIME(20000000); loop();
    ADVANCE_TIME(20000000); loop();
    ADVANCE_TIME(20000000); loop();
    ADVANCE_TIME(20000000); loop();
    ADVANCE_TIME(20000000); loop();
    ADVANCE_TIME(20000000); loop();
    ADVANCE_TIME(20000000); loop();
    ADVANCE_TIME(20000000); loop();
    ADVANCE_TIME(20000000); loop();
    ADVANCE_TIME(20000000); loop();
    ADVANCE_TIME(20000000); loop();
    ADVANCE_TIME(20000000); loop();
    ADVANCE_TIME(20000000); loop();
    ADVANCE_TIME(20000000); loop();
    ADVANCE_TIME(20000000); loop();
    ADVANCE_TIME(20000000); loop();
    ADVANCE_TIME(20000000); loop();
    ADVANCE_TIME(20000000); loop();
    ADVANCE_TIME(20000000); loop();
    ADVANCE_TIME(20000000); loop();
    ADVANCE_TIME(20000000); loop();
    ADVANCE_TIME(20000000); loop();
    ADVANCE_TIME(20000000); loop();
    ADVANCE_TIME(20000000); loop();
    ADVANCE_TIME(20000000); loop();
    ADVANCE_TIME(20000000); loop();
    ADVANCE_TIME(20000000); loop();
    ADVANCE_TIME(20000000); loop();
    ADVANCE_TIME(20000000); loop();
    ADVANCE_TIME(20000000); loop();
    ADVANCE_TIME(20000000); loop();
    ADVANCE_TIME(20000000); loop();
    ADVANCE_TIME(20000000); loop();
    ADVANCE_TIME(20000000); loop();
    ADVANCE_TIME(20000000); loop();
    ADVANCE_TIME(20000000); loop();
    ADVANCE_TIME(20000000); loop();
    ADVANCE_TIME(20000000); loop();
    ADVANCE_TIME(20000000); loop();
    ADVANCE_TIME(20000000); loop();
    ADVANCE_TIME(20000000); loop();
    ADVANCE_TIME(20000000); loop();
    ADVANCE_TIME(20000000); loop();
    ADVANCE_TIME(20000000); loop();
    ADVANCE_TIME(20000000); loop();
    ADVANCE_TIME(20000000); loop();
    ADVANCE_TIME(20000000); loop();
    ADVANCE_TIME(20000000); loop();
    ADVANCE_TIME(20000000); loop();
    ADVANCE_TIME(20000000); loop();
    ADVANCE_TIME(20000000); loop();
    ADVANCE_TIME(20000000); loop();
    ADVANCE_TIME(20000000); loop();
    ADVANCE_TIME(20000000); loop();
    ADVANCE_TIME(20000000); loop();
    ADVANCE_TIME(20000000); loop();
    ADVANCE_TIME(20000000); loop();
    ADVANCE_TIME(20000000); loop();
    ADVANCE_TIME(20000000); loop();
    ADVANCE_TIME(20000000); loop();
    ADVANCE_TIME(20000000); loop();
    ADVANCE_TIME(20000000); loop();
    ADVANCE_TIME(20000000); loop();
    ADVANCE_TIME(20000000); loop();
    ADVANCE_TIME(20000000); loop();
    ADVANCE_TIME(20000000); loop();
    ADVANCE_TIME(20000000); loop();
    ADVANCE_TIME(20000000); loop();
    ADVANCE_TIME(20000000); loop();
    ADVANCE_TIME(20000000); loop();
    ADVANCE_TIME(20000000); loop();
    ADVANCE_TIME(20000000); loop();
    ADVANCE_TIME(20000000); loop();
    ADVANCE_TIME(20000000); loop();
    ADVANCE_TIME(20000000); loop();
    ADVANCE_TIME(20000000); loop();
    ADVANCE_TIME(20000000); loop();
    ADVANCE_TIME(20000000); loop();
    ADVANCE_TIME(20000000); loop();
    ADVANCE_TIME(20000000); loop();
    ADVANCE_TIME(20000000); loop();
    ADVANCE_TIME(20000000); loop();
    ADVANCE_TIME(20000000); loop();
    ADVANCE_TIME(20000000); loop();
    ADVANCE_TIME(20000000); loop();
    ADVANCE_TIME(20000000); loop();
    ADVANCE_TIME(20000000); loop();
    ADVANCE_TIME(20000000); loop();
    ADVANCE_TIME(20000000); loop();
    ADVANCE_TIME(20000000); loop();
    ADVANCE_TIME(20000000); loop();
    ADVANCE_TIME(20000000); loop();
    ADVANCE_TIME(20000000); loop();
    ADVANCE_TIME(20000000); loop();
    ADVANCE_TIME(20000000); loop();
    ADVANCE_TIME(20000000); loop();
    ADVANCE_TIME(20000000); loop();
    ADVANCE_TIME(20000000); loop();
    ADVANCE_TIME(20000000); loop();
    ADVANCE_TIME(20000000); loop();
    ADVANCE_TIME(20000000); loop();
    ADVANCE_TIME(20000000); loop();
    ADVANCE_TIME(20000000); loop();
    ADVANCE_TIME(20000000); loop();
    ADVANCE_TIME(20000000); loop();
    ADVANCE_TIME(20000000); loop();
    ADVANCE_TIME(20000000); loop();
    ADVANCE_TIME(20000000); loop();
    ADVANCE_TIME(20000000); loop();
    ADVANCE_TIME(20000000); loop();
    ADVANCE_TIME(20000000); loop();
    ADVANCE_TIME(20000000); loop();
    ADVANCE_TIME(20000000); loop();
    ADVANCE_TIME(20000000); loop();
    ADVANCE_TIME(20000000); loop();
    ADVANCE_TIME(20000000); loop();
    ADVANCE_TIME(20000000); loop();
    ADVANCE_TIME(20000000); loop();
    ADVANCE_TIME(20000000); loop();
    ADVANCE_TIME(20000000); loop();
    ADVANCE_TIME(20000000); loop();
    ADVANCE_TIME(20000000); loop();
    ADVANCE_TIME(20000000); loop();
    ADVANCE_TIME(20000000); loop();
    ADVANCE_TIME(20000000); loop();
    ADVANCE_TIME(20000000); loop();
    ADVANCE_TIME(20000000); loop();
    ADVANCE_TIME(20000000); loop();
    ADVANCE_TIME(20000000); loop();
    ADVANCE_TIME(20000000); loop();
    ADVANCE_TIME(20000000); loop();
    ADVANCE_TIME(20000000); loop();
    ADVANCE_TIME(20000000); loop();
    ADVANCE_TIME(20000000); loop();
    ADVANCE_TIME(20000000); loop();
    ADVANCE_TIME(20000000); loop();
    ADVANCE_TIME(20000000); loop();
    ADVANCE_TIME(20000000); loop();
    ADVANCE_TIME(20000000); loop();
    ADVANCE_TIME(20000000); loop();
    ADVANCE_TIME(20000000); loop();
    ADVANCE_TIME(20000000); loop();
    ADVANCE_TIME(20000000); loop();
    ADVANCE_TIME(20000000); loop();
    ADVANCE_TIME(20000000); loop();
    ADVANCE_TIME(20000000); loop();
    ADVANCE_TIME(20000000); loop();
    ADVANCE_TIME(20000000); loop();
    ADVANCE_TIME(20000000); loop();
    ADVANCE_TIME(20000000); loop();
    ADVANCE_TIME(20000000); loop();
    ADVANCE_TIME(20000000); loop();
    ADVANCE_TIME(20000000); loop();
    ADVANCE_TIME(20000000); loop();
    ADVANCE_TIME(20000000); loop();
    ADVANCE_TIME(20000000); loop();
    ADVANCE_TIME(20000000); loop();
    ADVANCE_TIME(20000000); loop();
    ADVANCE_TIME(20000000); loop();
    ADVANCE_TIME(20000000); loop();
    ADVANCE_TIME(20000000); loop();
    ADVANCE_TIME(20000000); loop();
    ADVANCE_TIME(20000000); loop();
    ADVANCE_TIME(20000000); loop();
    ADVANCE_TIME(20000000); loop();
    ADVANCE_TIME(20000000); loop();
    ADVANCE_TIME(20000000); loop();
    ADVANCE_TIME(20000000); loop();
    ADVANCE_TIME(20000000); loop();
    ADVANCE_TIME(20000000); loop();
    ADVANCE_TIME(20000000); loop();
    ADVANCE_TIME(20000000); loop();
    ADVANCE_TIME(20000000); loop();
    ADVANCE_TIME(20000000); loop();
    ADVANCE_TIME(20000000); loop();
    ADVANCE_TIME(20000000); loop();
    ADVANCE_TIME(20000000); loop();
    ADVANCE_TIME(20000000); loop();
    ADVANCE_TIME(20000000); loop();
    ADVANCE_TIME(20000000); loop();
    ADVANCE_TIME(20000000); loop();
    ADVANCE_TIME(20000000); loop();
    ADVANCE_TIME(20000000); loop();
    ADVANCE_TIME(20000000); loop();
    ADVANCE_TIME(20000000); loop();
    ADVANCE_TIME(20000000); loop();
    ADVANCE_TIME(20000000); loop();
    ADVANCE_TIME(20000000); loop();
    ADVANCE_TIME(20000000); loop();
    ADVANCE_TIME(20000000); loop();
    ADVANCE_TIME(20000000); loop();
    ADVANCE_TIME(20000000); loop();
    ADVANCE_TIME(20000000); loop();
    ADVANCE_TIME(20000000); loop();
    ADVANCE_TIME(20000000); loop();
    ADVANCE_TIME(20000000); loop();
    ADVANCE_TIME(20000000); loop();
    ADVANCE_TIME(20000000); loop();
    ADVANCE_TIME(20000000); loop();
    ADVANCE_TIME(20000000); loop();
    ADVANCE_TIME(20000000); loop();
    ADVANCE_TIME(20000000); loop();
    ADVANCE_TIME(20000000); loop();
    ADVANCE_TIME(20000000); loop();
    ADVANCE_TIME(20000000); loop();
    ADVANCE_TIME(20000000); loop();
    ADVANCE_TIME(20000000); loop();
    ADVANCE_TIME(20000000); loop();
    ADVANCE_TIME(20000000); loop();
    ADVANCE_TIME(20000000); loop();
    ADVANCE_TIME(20000000); loop();
    ADVANCE_TIME(20000000); loop();
    ADVANCE_TIME(20000000); loop();
    ADVANCE_TIME(20000000); loop();
    ADVANCE_TIME(20000000); loop();
    ADVANCE_TIME(20000000); loop();
    ADVANCE_TIME(20000000); loop();
    ADVANCE_TIME(20000000); loop();
    ADVANCE_TIME(20000000); loop();
    ADVANCE_TIME(20000000); loop();
    ADVANCE_TIME(20000000); loop();
    ADVANCE_TIME(20000000); loop();
    ADVANCE_TIME(20000000); loop();
    ADVANCE_TIME(20000000); loop();
    ADVANCE_TIME(20000000); loop();
    ADVANCE_TIME(20000000); loop();
    ADVANCE_TIME(20000000); loop();
    ADVANCE_TIME(20000000); loop();
    ADVANCE_TIME(20000000); loop();
    ADVANCE_TIME(20000000); loop();
    ADVANCE_TIME(20000000); loop();
    ADVANCE_TIME(20000000); loop();
    ADVANCE_TIME(20000000); loop();
    ADVANCE_TIME(20000000); loop();
    ADVANCE_TIME(20000000); loop();
    ADVANCE_TIME(20000000); loop();
    ADVANCE_TIME(20000000); loop();
    ADVANCE_TIME(20000000); loop();
    ADVANCE_TIME(20000000); loop();
    ADVANCE_TIME(20000000); loop();
    ADVANCE_TIME(20000000); loop();
    ADVANCE_TIME(20000000); loop();
    ADVANCE_TIME(20000000); loop();
    ADVANCE_TIME(20000000); loop();
    ADVANCE_TIME(20000000); loop();
    ADVANCE_TIME(20000000); loop();
    ADVANCE_TIME(20000000); loop();
    ADVANCE_TIME(20000000); loop();
    ADVANCE_TIME(20000000); loop();
    ADVANCE_TIME(20000000); loop();
    ADVANCE_TIME(20000000); loop();
    ADVANCE_TIME(20000000); loop();
    ADVANCE_TIME(20000000); loop();
    ADVANCE_TIME(20000000); loop();
    ADVANCE_TIME(20000000); loop();
    ADVANCE_TIME(20000000); loop();
    ADVANCE_TIME(20000000); loop();
    ADVANCE_TIME(20000000); loop();
    ADVANCE_TIME(20000000); loop();
    ADVANCE_TIME(20000000); loop();
    ADVANCE_TIME(20000000); loop();
    ADVANCE_TIME(20000000); loop();
    ADVANCE_TIME(20000000); loop();
    ADVANCE_TIME(20000000); loop();
    ADVANCE_TIME(20000000); loop();
    ADVANCE_TIME(20000000); loop();
    ADVANCE_TIME(20000000); loop();
    ADVANCE_TIME(20000000); loop();
    ADVANCE_TIME(20000000); loop();
    ADVANCE_TIME(20000000); loop();
    ADVANCE_TIME(20000000); loop();
    ADVANCE_TIME(20000000); loop();
    ADVANCE_TIME(20000000); loop();
    ADVANCE_TIME(20000000); loop();
    ADVANCE_TIME(20000000); loop();
    ADVANCE_TIME(20000000); loop();
    ADVANCE_TIME(20000000); loop();
    ADVANCE_TIME(20000000); loop();
    ADVANCE_TIME(20000000); loop();
    ADVANCE_TIME(20000000); loop();
    ADVANCE_TIME(20000000); loop();
    ADVANCE_TIME(20000000); loop();
    ADVANCE_TIME(20000000); loop();
    ADVANCE_TIME(20000000); loop();
    ADVANCE_TIME(20000000); loop();
    ADVANCE_TIME(20000000); loop();
    ADVANCE_TIME(20000000); loop();
    ADVANCE_TIME(20000000); loop();
    ADVANCE_TIME(20000000); loop();
    ADVANCE_TIME(20000000); loop();
    ADVANCE_TIME(20000000); loop();
    ADVANCE_TIME(20000000); loop();
    ADVANCE_TIME(20000000); loop();
    ADVANCE_TIME(20000000); loop();
    ADVANCE_TIME(20000000); loop();
    ADVANCE_TIME(20000000); loop();
    ADVANCE_TIME(20000000); loop();
    ADVANCE_TIME(20000000); loop();
    ADVANCE_TIME(20000000); loop();
    ADVANCE_TIME(20000000); loop();
    ADVANCE_TIME(20000000); loop();
    ADVANCE_TIME(20000000); loop();
    ADVANCE_TIME(20000000); loop();
    ADVANCE_TIME(20000000); loop();
    ADVANCE_TIME(20000000); loop();
    ADVANCE_TIME(20000000); loop();
    ADVANCE_TIME(20000000); loop();
    ADVANCE_TIME(20000000); loop();
    ADVANCE_TIME(20000000); loop();
    ADVANCE_TIME(20000000); loop();
    ADVANCE_TIME(20000000); loop();
    ADVANCE_TIME(20000000); loop();
    ADVANCE_TIME(20000000); loop();
    ADVANCE_TIME(20000000); loop();
    ADVANCE_TIME(20000000); loop();
    ADVANCE_TIME(20000000); loop();
    ADVANCE_TIME(20000000); loop();
    ADVANCE_TIME(20000000); loop();
    ADVANCE_TIME(20000000); loop();
    ADVANCE_TIME(20000000); loop();
    ADVANCE_TIME(20000000); loop();
    ADVANCE_TIME(20000000); loop();
    ADVANCE_TIME(20000000); loop();
    ADVANCE_TIME(20000000); loop();
    ADVANCE_TIME(20000000); loop();
    ADVANCE_TIME(20000000); loop();
    ADVANCE_TIME(20000000); loop();
    ADVANCE_TIME(20000000); loop();
    ADVANCE_TIME(20000000); loop();
    ADVANCE_TIME(20000000); loop();
    ADVANCE_TIME(20000000); loop();
    ADVANCE_TIME(20000000); loop();
    ADVANCE_TIME(20000000); loop();
    ADVANCE_TIME(20000000); loop();
    ADVANCE_TIME(20000000); loop();
    ADVANCE_TIME(20000000); loop();
    ADVANCE_TIME(20000000); loop();
    ADVANCE_TIME(20000000); loop();
    ADVANCE_TIME(20000000); loop();
    ADVANCE_TIME(20000000); loop();
    ADVANCE_TIME(20000000); loop();
    ADVANCE_TIME(20000000); loop();
    ADVANCE_TIME(20000000); loop();
    ADVANCE_TIME(20000000); loop();
    ADVANCE_TIME(20000000); loop();
    ADVANCE_TIME(20000000); loop();
    ADVANCE_TIME(20000000); loop();
    ADVANCE_TIME(20000000); loop();
    ADVANCE_TIME(20000000); loop();
    ADVANCE_TIME(20000000); loop();
    ADVANCE_TIME(20000000); loop();
    ADVANCE_TIME(20000000); loop();
    ADVANCE_TIME(20000000); loop();
    ADVANCE_TIME(20000000); loop();
    ADVANCE_TIME(20000000); loop();
    ADVANCE_TIME(20000000); loop();
    ADVANCE_TIME(20000000); loop();
    ADVANCE_TIME(20000000); loop();
    ADVANCE_TIME(20000000); loop();
    ADVANCE_TIME(20000000); loop();
    ADVANCE_TIME(20000000); loop();
    ADVANCE_TIME(20000000); loop();
    ADVANCE_TIME(20000000); loop();
    ADVANCE_TIME(20000000); loop();
    ADVANCE_TIME(20000000); loop();
    ADVANCE_TIME(20000000); loop();
    ADVANCE_TIME(20000000); loop();
    ADVANCE_TIME(20000000); loop();
    ADVANCE_TIME(20000000); loop();
    ADVANCE_TIME(20000000); loop();
    ADVANCE_TIME(20000000); loop();
    ADVANCE_TIME(20000000); loop();
    ADVANCE_TIME(20000000); loop();
    ADVANCE_TIME(20000000); loop();
    ADVANCE_TIME(20000000); loop();
    ADVANCE_TIME(20000000); loop();
    ADVANCE_TIME(20000000); loop();
    ADVANCE_TIME(20000000); loop();
    ADVANCE_TIME(20000000); loop();
    ADVANCE_TIME(20000000); loop();
    ADVANCE_TIME(20000000); loop();
    ADVANCE_TIME(20000000); loop();
    ADVANCE_TIME(20000000); loop();
    ADVANCE_TIME(20000000); loop();
    ADVANCE_TIME(20000000); loop();
    ADVANCE_TIME(20000000); loop();
    ADVANCE_TIME(20000000); loop();
    ADVANCE_TIME(20000000); loop();
    ADVANCE_TIME(20000000); loop();
    ADVANCE_TIME(20000000); loop();
    ADVANCE_TIME(20000000); loop();
    ADVANCE_TIME(20000000); loop();
    ADVANCE_TIME(20000000); loop();
    ADVANCE_TIME(20000000); loop();
    ADVANCE_TIME(20000000); loop();
    ADVANCE_TIME(20000000); loop();
    ADVANCE_TIME(20000000); loop();
    ADVANCE_TIME(20000000); loop();
    ADVANCE_TIME(20000000); loop();
    ADVANCE_TIME(20000000); loop();
    ADVANCE_TIME(20000000); loop();
    ADVANCE_TIME(20000000); loop();
    ADVANCE_TIME(20000000); loop();
    ADVANCE_TIME(20000000); loop();
    ADVANCE_TIME(20000000); loop();
    ADVANCE_TIME(20000000); loop();
    ADVANCE_TIME(20000000); loop();
    ADVANCE_TIME(20000000); loop();
    ADVANCE_TIME(20000000); loop();
    ADVANCE_TIME(20000000); loop();
    ADVANCE_TIME(20000000); loop();
    ADVANCE_TIME(20000000); loop();
    ADVANCE_TIME(20000000); loop();
    ADVANCE_TIME(20000000); loop();
    ADVANCE_TIME(20000000); loop();
    ADVANCE_TIME(20000000); loop();
    ADVANCE_TIME(20000000); loop();
    ADVANCE_TIME(20000000); loop();
    ADVANCE_TIME(20000000); loop();
    ADVANCE_TIME(20000000); loop();
    ADVANCE_TIME(20000000); loop();
    ADVANCE_TIME(20000000); loop();
    ADVANCE_TIME(20000000); loop();
    ADVANCE_TIME(20000000); loop();
    ADVANCE_TIME(20000000); loop();
    ADVANCE_TIME(20000000); loop();
    ADVANCE_TIME(20000000); loop();
    ADVANCE_TIME(20000000); loop();
    ADVANCE_TIME(20000000); loop();
    ADVANCE_TIME(20000000); loop();
    ADVANCE_TIME(20000000); loop();
    ADVANCE_TIME(20000000); loop();
    ADVANCE_TIME(20000000); loop();
    ADVANCE_TIME(20000000); loop();
    ADVANCE_TIME(20000000); loop();
    ADVANCE_TIME(20000000); loop();
    ADVANCE_TIME(20000000); loop();
    ADVANCE_TIME(20000000); loop();
    ADVANCE_TIME(20000000); loop();
    ADVANCE_TIME(20000000); loop();
    ADVANCE_TIME(20000000); loop();
    ADVANCE_TIME(20000000); loop();
    ADVANCE_TIME(20000000); loop();
    ADVANCE_TIME(20000000); loop();
    ADVANCE_TIME(20000000); loop();
    ADVANCE_TIME(20000000); loop();
    ADVANCE_TIME(20000000); loop();
    ADVANCE_TIME(20000000); loop();
    ADVANCE_TIME(20000000); loop();
    ADVANCE_TIME(20000000); loop();
    ADVANCE_TIME(20000000); loop();
    ADVANCE_TIME(20000000); loop();
    ADVANCE_TIME(20000000); loop();
    ADVANCE_TIME(20000000); loop();
    ADVANCE_TIME(20000000); loop();
    ADVANCE_TIME(20000000); loop();
    ADVANCE_TIME(20000000); loop();
    ADVANCE_TIME(20000000); loop();
    ADVANCE_TIME(20000000); loop();
    ADVANCE_TIME(20000000); loop();
    ADVANCE_TIME(20000000); loop();
    ADVANCE_TIME(20000000); loop();
    ADVANCE_TIME(20000000); loop();
    ADVANCE_TIME(20000000); loop();
    ADVANCE_TIME(20000000); loop();
    ADVANCE_TIME(20000000); loop();
    ADVANCE_TIME(20000000); loop();
    ADVANCE_TIME(20000000); loop();
    ADVANCE_TIME(20000000); loop();
    ADVANCE_TIME(20000000); loop();
    ADVANCE_TIME(20000000); loop();
    ADVANCE_TIME(20000000); loop();
    ADVANCE_TIME(20000000); loop();
    ADVANCE_TIME(20000000); loop();
    ADVANCE_TIME(20000000); loop();
    ADVANCE_TIME(20000000); loop();
    ADVANCE_TIME(20000000); loop();
    ADVANCE_TIME(20000000); loop();
    ADVANCE_TIME(20000000); loop();
    ADVANCE_TIME(20000000); loop();
    ADVANCE_TIME(20000000); loop();
    ADVANCE_TIME(20000000); loop();
    ADVANCE_TIME(20000000); loop();
    ADVANCE_TIME(20000000); loop();
    ADVANCE_TIME(20000000); loop();
    ADVANCE_TIME(20000000); loop();
    ADVANCE_TIME(20000000); loop();
    ADVANCE_TIME(20000000); loop();
    ADVANCE_TIME(20000000); loop();
    ADVANCE_TIME(20000000); loop();
    ADVANCE_TIME(20000000); loop();
    ADVANCE_TIME(20000000); loop();
    ADVANCE_TIME(20000000); loop();
    ADVANCE_TIME(20000000); loop();
    ADVANCE_TIME(20000000); loop();
    ADVANCE_TIME(20000000); loop();
    ADVANCE_TIME(20000000); loop();
    ADVANCE_TIME(20000000); loop();
    ADVANCE_TIME(20000000); loop();
    ADVANCE_TIME(20000000); loop();
    ADVANCE_TIME(20000000); loop();
    ADVANCE_TIME(20000000); loop();
    ADVANCE_TIME(20000000); loop();
    ADVANCE_TIME(20000000); loop();
    ADVANCE_TIME(20000000); loop();
    ADVANCE_TIME(20000000); loop();
    ADVANCE_TIME(20000000); loop();
    ADVANCE_TIME(20000000); loop();
    ADVANCE_TIME(20000000); loop();
    ADVANCE_TIME(20000000); loop();
    ADVANCE_TIME(20000000); loop();
    ADVANCE_TIME(20000000); loop();
    ADVANCE_TIME(20000000); loop();
    ADVANCE_TIME(20000000); loop();
    ADVANCE_TIME(20000000); loop();
    ADVANCE_TIME(20000000); loop();
    ADVANCE_TIME(20000000); loop();
    ADVANCE_TIME(20000000); loop();
    ADVANCE_TIME(20000000); loop();
    ADVANCE_TIME(20000000); loop();
    ADVANCE_TIME(20000000); loop();
    ADVANCE_TIME(20000000); loop();
    ADVANCE_TIME(20000000); loop();
    ADVANCE_TIME(20000000); loop();
    ADVANCE_TIME(20000000); loop();
    ADVANCE_TIME(20000000); loop();
    ADVANCE_TIME(20000000); loop();
    ADVANCE_TIME(20000000); loop();
    ADVANCE_TIME(20000000); loop();
    ADVANCE_TIME(20000000); loop();
    ADVANCE_TIME(20000000); loop();
    ADVANCE_TIME(20000000); loop();
    ADVANCE_TIME(20000000); loop();
    ADVANCE_TIME(20000000); loop();
    ADVANCE_TIME(20000000); loop();
    ADVANCE_TIME(20000000); loop();
    ADVANCE_TIME(20000000); loop();
    ADVANCE_TIME(20000000); loop();
    ADVANCE_TIME(20000000); loop();
    ADVANCE_TIME(20000000); loop();
    ADVANCE_TIME(20000000); loop();
    ADVANCE_TIME(20000000); loop();
    ADVANCE_TIME(20000000); loop();
    ADVANCE_TIME(20000000); loop();
    ADVANCE_TIME(20000000); loop();
    ADVANCE_TIME(20000000); loop();
    ADVANCE_TIME(20000000); loop();
    ADVANCE_TIME(20000000); loop();
    ADVANCE_TIME(20000000); loop();
    ADVANCE_TIME(20000000); loop();
    ADVANCE_TIME(20000000); loop();
    ADVANCE_TIME(20000000); loop();
    ADVANCE_TIME(20000000); loop();
    ADVANCE_TIME(20000000); loop();
    ADVANCE_TIME(20000000); loop();
    ADVANCE_TIME(20000000); loop();
    ADVANCE_TIME(20000000); loop();
    ADVANCE_TIME(20000000); loop();
    ADVANCE_TIME(20000000); loop();
    ADVANCE_TIME(20000000); loop();
    ADVANCE_TIME(20000000); loop();
    ADVANCE_TIME(20000000); loop();
    ADVANCE_TIME(20000000); loop();
    ADVANCE_TIME(20000000); loop();
    ADVANCE_TIME(20000000); loop();
    ADVANCE_TIME(20000000); loop();
    ADVANCE_TIME(20000000); loop();
    ADVANCE_TIME(20000000); loop();
    ADVANCE_TIME(20000000); loop();
    ADVANCE_TIME(20000000); loop();
    ADVANCE_TIME(20000000); loop();
    ADVANCE_TIME(20000000); loop();
    ADVANCE_TIME(20000000); loop();
    ADVANCE_TIME(20000000); loop();
    ADVANCE_TIME(20000000); loop();
    ADVANCE_TIME(20000000); loop();
    ADVANCE_TIME(20000000); loop();
    ADVANCE_TIME(20000000); loop();
    ADVANCE_TIME(20000000); loop();
    ADVANCE_TIME(20000000); loop();
    ADVANCE_TIME(20000000); loop();
    ADVANCE_TIME(20000000); loop();
    ADVANCE_TIME(20000000); loop();
    ADVANCE_TIME(20000000); loop();
    ADVANCE_TIME(20000000); loop();
    ADVANCE_TIME(20000000); loop();
    ADVANCE_TIME(20000000); loop();
    ADVANCE_TIME(20000000); loop();
    ADVANCE_TIME(20000000); loop();
    ADVANCE_TIME(20000000); loop();
    ADVANCE_TIME(20000000); loop();
    ADVANCE_TIME(20000000); loop();
    ADVANCE_TIME(20000000); loop();
    ADVANCE_TIME(20000000); loop();
    ADVANCE_TIME(20000000); loop();
    ADVANCE_TIME(20000000); loop();
    ADVANCE_TIME(20000000); loop();
    ADVANCE_TIME(20000000); loop();
    ADVANCE_TIME(20000000); loop();
    ADVANCE_TIME(20000000); loop();
    ADVANCE_TIME(20000000); loop();
    ADVANCE_TIME(20000000); loop();
    ADVANCE_TIME(20000000); loop();
    ADVANCE_TIME(20000000); loop();
    ADVANCE_TIME(20000000); loop();
    ADVANCE_TIME(20000000); loop();
    ADVANCE_TIME(20000000); loop();
    ADVANCE_TIME(20000000); loop();
    ADVANCE_TIME(20000000); loop();
    ADVANCE_TIME(20000000); loop();
    ADVANCE_TIME(20000000); loop();
    ADVANCE_TIME(20000000); loop();
    ADVANCE_TIME(20000000); loop();
    ADVANCE_TIME(20000000); loop();
    ADVANCE_TIME(20000000); loop();
    ADVANCE_TIME(20000000); loop();
    ADVANCE_TIME(20000000); loop();
    ADVANCE_TIME(20000000); loop();
    ADVANCE_TIME(20000000); loop();
    ADVANCE_TIME(20000000); loop();
    ADVANCE_TIME(20000000); loop();
    ADVANCE_TIME(20000000); loop();
    ADVANCE_TIME(20000000); loop();
    ADVANCE_TIME(20000000); loop();
    ADVANCE_TIME(20000000); loop();
    ADVANCE_TIME(20000000); loop();
    ADVANCE_TIME(20000000); loop();
    ADVANCE_TIME(20000000); loop();
    ADVANCE_TIME(20000000); loop();
    ADVANCE_TIME(20000000); loop();
    ADVANCE_TIME(20000000); loop();
    ADVANCE_TIME(20000000); loop();
    ADVANCE_TIME(20000000); loop();
    ADVANCE_TIME(20000000); loop();
    ADVANCE_TIME(20000000); loop();
    ADVANCE_TIME(20000000); loop();
    ADVANCE_TIME(20000000); loop();
    ADVANCE_TIME(20000000); loop();
    ADVANCE_TIME(20000000); loop();
    ADVANCE_TIME(20000000); loop();
    ADVANCE_TIME(20000000); loop();
    ADVANCE_TIME(20000000); loop();
    ADVANCE_TIME(20000000); loop();
    ADVANCE_TIME(20000000); loop();
    ADVANCE_TIME(20000000); loop();
    ADVANCE_TIME(20000000); loop();
    ADVANCE_TIME(20000000); loop();
    ADVANCE_TIME(20000000); loop();
    ADVANCE_TIME(20000000); loop();
    ADVANCE_TIME(20000000); loop();
    ADVANCE_TIME(20000000); loop();
    ADVANCE_TIME(20000000); loop();
    ADVANCE_TIME(20000000); loop();
    ADVANCE_TIME(20000000); loop();
    ADVANCE_TIME(20000000); loop();
    ADVANCE_TIME(20000000); loop();
    ADVANCE_TIME(20000000); loop();
    ADVANCE_TIME(20000000); loop();
    ADVANCE_TIME(20000000); loop();
    ADVANCE_TIME(20000000); loop();
    ADVANCE_TIME(20000000); loop();
    ADVANCE_TIME(20000000); loop();
    ADVANCE_TIME(20000000); loop();
    ADVANCE_TIME(20000000); loop();
    ADVANCE_TIME(20000000); loop();
    ADVANCE_TIME(20000000); loop();
    ADVANCE_TIME(20000000); loop();
    ADVANCE_TIME(20000000); loop();
    ADVANCE_TIME(20000000); loop();
    ADVANCE_TIME(20000000); loop();
    ADVANCE_TIME(20000000); loop();
    ADVANCE_TIME(20000000); loop();
    ADVANCE_TIME(20000000); loop();
    ADVANCE_TIME(20000000); loop();
    ADVANCE_TIME(20000000); loop();
    ADVANCE_TIME(20000000); loop();
    ADVANCE_TIME(20000000); loop();
    ADVANCE_TIME(20000000); loop();
    ADVANCE_TIME(20000000); loop();
    ADVANCE_TIME(20000000); loop();
    ADVANCE_TIME(20000000); loop();
    ADVANCE_TIME(20000000); loop();
    ADVANCE_TIME(20000000); loop();
    ADVANCE_TIME(20000000); loop();
    ADVANCE_TIME(20000000); loop();
    ADVANCE_TIME(20000000); loop();
    ADVANCE_TIME(20000000); loop();
    ADVANCE_TIME(20000000); loop();
    ADVANCE_TIME(20000000); loop();
    ADVANCE_TIME(20000000); loop();
    ADVANCE_TIME(20000000); loop();
    ADVANCE_TIME(20000000); loop();
    ADVANCE_TIME(20000000); loop();
    ADVANCE_TIME(20000000); loop();
    ADVANCE_TIME(20000000); loop();
    ADVANCE_TIME(20000000); loop();
    ADVANCE_TIME(20000000); loop();
    ADVANCE_TIME(20000000); loop();
    ADVANCE_TIME(20000000); loop();
    ADVANCE_TIME(20000000); loop();
    ADVANCE_TIME(20000000); loop();
    ADVANCE_TIME(20000000); loop();
    ADVANCE_TIME(20000000); loop();
    ADVANCE_TIME(20000000); loop();
    ADVANCE_TIME(20000000); loop();
    ADVANCE_TIME(20000000); loop();
    ADVANCE_TIME(20000000); loop();
    ADVANCE_TIME(20000000); loop();
    ADVANCE_TIME(20000000); loop();
    ADVANCE_TIME(20000000); loop();
    ADVANCE_TIME(20000000); loop();
    ADVANCE_TIME(20000000); loop();
    ADVANCE_TIME(20000000); loop();
    ADVANCE_TIME(20000000); loop();
    ADVANCE_TIME(20000000); loop();
    ADVANCE_TIME(20000000); loop();
    ADVANCE_TIME(20000000); loop();
    ADVANCE_TIME(20000000); loop();
    ADVANCE_TIME(20000000); loop();
    ADVANCE_TIME(20000000); loop();
    ADVANCE_TIME(20000000); loop();
    ADVANCE_TIME(20000000); loop();
    ADVANCE_TIME(20000000); loop();
    ADVANCE_TIME(20000000); loop();
    ADVANCE_TIME(20000000); loop();
    ADVANCE_TIME(20000000); loop();
    ADVANCE_TIME(20000000); loop();
    ADVANCE_TIME(20000000); loop();
    ADVANCE_TIME(20000000); loop();
    ADVANCE_TIME(20000000); loop();
    ADVANCE_TIME(20000000); loop();
    ADVANCE_TIME(20000000); loop();
    ADVANCE_TIME(20000000); loop();
    ADVANCE_TIME(20000000); loop();
    ADVANCE_TIME(20000000); loop();
    ADVANCE_TIME(20000000); loop();
    ADVANCE_TIME(20000000); loop();
    ADVANCE_TIME(20000000); loop();
    ADVANCE_TIME(20000000); loop();
    ADVANCE_TIME(20000000); loop();
    ADVANCE_TIME(20000000); loop();
    ADVANCE_TIME(20000000); loop();
    ADVANCE_TIME(20000000); loop();
    ADVANCE_TIME(20000000); loop();
    ADVANCE_TIME(20000000); loop();
    ADVANCE_TIME(20000000); loop();
    ADVANCE_TIME(20000000); loop();
    ADVANCE_TIME(20000000); loop();
    ADVANCE_TIME(20000000); loop();
    ADVANCE_TIME(20000000); loop();
    ADVANCE_TIME(20000000); loop();
    ADVANCE_TIME(20000000); loop();
    ADVANCE_TIME(20000000); loop();
    ADVANCE_TIME(20000000); loop();
    ADVANCE_TIME(20000000); loop();
    ADVANCE_TIME(20000000); loop();
    ADVANCE_TIME(20000000); loop();
    ADVANCE_TIME(20000000); loop();
    ADVANCE_TIME(20000000); loop();
    ADVANCE_TIME(20000000); loop();
    ADVANCE_TIME(20000000); loop();
    ADVANCE_TIME(20000000); loop();
    ADVANCE_TIME(20000000); loop();
    ADVANCE_TIME(20000000); loop();
    ADVANCE_TIME(20000000); loop();
    ADVANCE_TIME(20000000); loop();
    ADVANCE_TIME(20000000); loop();
    ADVANCE_TIME(20000000); loop();
    ADVANCE_TIME(20000000); loop();
    ADVANCE_TIME(20000000); loop();
    ADVANCE_TIME(20000000); loop();
    ADVANCE_TIME(20000000); loop();
    ADVANCE_TIME(20000000); loop();
    ADVANCE_TIME(20000000); loop();
    ADVANCE_TIME(20000000); loop();
    ADVANCE_TIME(20000000); loop();
    ADVANCE_TIME(20000000); loop();
    ADVANCE_TIME(20000000); loop();
    ADVANCE_TIME(20000000); loop();
    ADVANCE_TIME(20000000); loop();
    ADVANCE_TIME(20000000); loop();
    ADVANCE_TIME(20000000); loop();
    ADVANCE_TIME(20000000); loop();
    ADVANCE_TIME(20000000); loop();
    ADVANCE_TIME(20000000); loop();
    ADVANCE_TIME(20000000); loop();
    ADVANCE_TIME(20000000); loop();
    ADVANCE_TIME(20000000); loop();
    ADVANCE_TIME(20000000); loop();
    ADVANCE_TIME(20000000); loop();
    ADVANCE_TIME(20000000); loop();
    ADVANCE_TIME(20000000); loop();
    ADVANCE_TIME(20000000); loop();
    ADVANCE_TIME(20000000); loop();
    ADVANCE_TIME(20000000); loop();
    ADVANCE_TIME(20000000); loop();
    ADVANCE_TIME(20000000); loop();
    ADVANCE_TIME(20000000); loop();
    ADVANCE_TIME(20000000); loop();
    ADVANCE_TIME(20000000); loop();
    ADVANCE_TIME(20000000); loop();
    ADVANCE_TIME(20000000); loop();
    ADVANCE_TIME(20000000); loop();
    ADVANCE_TIME(20000000); loop();
    ADVANCE_TIME(20000000); loop();
    ADVANCE_TIME(20000000); loop();
    ADVANCE_TIME(20000000); loop();
    ADVANCE_TIME(20000000); loop();
    ADVANCE_TIME(20000000); loop();
    ADVANCE_TIME(20000000); loop();
    ADVANCE_TIME(20000000); loop();
    ADVANCE_TIME(20000000); loop();
    ADVANCE_TIME(20000000); loop();
    ADVANCE_TIME(20000000); loop();
    ADVANCE_TIME(20000000); loop();
    ADVANCE_TIME(20000000); loop();
    ADVANCE_TIME(20000000); loop();
    ADVANCE_TIME(20000000); loop();
    ADVANCE_TIME(20000000); loop();
    ADVANCE_TIME(20000000); loop();
    ADVANCE_TIME(20000000); loop();
    ADVANCE_TIME(20000000); loop();
    ADVANCE_TIME(20000000); loop();
    ADVANCE_TIME(20000000); loop();
    ADVANCE_TIME(20000000); loop();
    ADVANCE_TIME(20000000); loop();
    ADVANCE_TIME(20000000); loop();
    ADVANCE_TIME(20000000); loop();
    ADVANCE_TIME(20000000); loop();
    ADVANCE_TIME(20000000); loop();
    ADVANCE_TIME(20000000); loop();
    ADVANCE_TIME(20000000); loop();
    ADVANCE_TIME(20000000); loop();
    ADVANCE_TIME(20000000); loop();
    ADVANCE_TIME(20000000); loop();
    ADVANCE_TIME(20000000); loop();
    ADVANCE_TIME(20000000); loop();
    ADVANCE_TIME(20000000); loop();
    ADVANCE_TIME(20000000); loop();
    ADVANCE_TIME(20000000); loop();
    ADVANCE_TIME(20000000); loop();
    ADVANCE_TIME(20000000); loop();
    ADVANCE_TIME(20000000); loop();
    ADVANCE_TIME(20000000); loop();
    ADVANCE_TIME(20000000); loop();
    ADVANCE_TIME(20000000); loop();
    ADVANCE_TIME(20000000); loop();
    ADVANCE_TIME(20000000); loop();
    ADVANCE_TIME(20000000); loop();
    ADVANCE_TIME(20000000); loop();
    ADVANCE_TIME(20000000); loop();
    ADVANCE_TIME(20000000); loop();
    ADVANCE_TIME(20000000); loop();
    ADVANCE_TIME(20000000); loop();
    ADVANCE_TIME(20000000); loop();
    ADVANCE_TIME(20000000); loop();
    ADVANCE_TIME(20000000); loop();
    ADVANCE_TIME(20000000); loop();
    ADVANCE_TIME(20000000); loop();
    ADVANCE_TIME(20000000); loop();
    ADVANCE_TIME(20000000); loop();
    ADVANCE_TIME(20000000); loop();
    ADVANCE_TIME(20000000); loop();
    ADVANCE_TIME(20000000); loop();
    ADVANCE_TIME(20000000); loop();
    ADVANCE_TIME(20000000); loop();
    ADVANCE_TIME(20000000); loop();
    ADVANCE_TIME(20000000); loop();
    ADVANCE_TIME(20000000); loop();
    ADVANCE_TIME(20000000); loop();
    ADVANCE_TIME(20000000); loop();
    ADVANCE_TIME(20000000); loop();
    ADVANCE_TIME(20000000); loop();
    ADVANCE_TIME(20000000); loop();
    ADVANCE_TIME(20000000); loop();
    ADVANCE_TIME(20000000); loop();
    ADVANCE_TIME(20000000); loop();
    ADVANCE_TIME(20000000); loop();
    ADVANCE_TIME(20000000); loop();
    ADVANCE_TIME(20000000); loop();
    ADVANCE_TIME(20000000); loop();
    ADVANCE_TIME(20000000); loop();
    ADVANCE_TIME(20000000); loop();
    ADVANCE_TIME(20000000); loop();
    ADVANCE_TIME(20000000); loop();
    ADVANCE_TIME(20000000); loop();
    ADVANCE_TIME(20000000); loop();
    ADVANCE_TIME(20000000); loop();
    ADVANCE_TIME(20000000); loop();
    ADVANCE_TIME(20000000); loop();
    ADVANCE_TIME(20000000); loop();
    ADVANCE_TIME(20000000); loop();
    ADVANCE_TIME(20000000); loop();
    ADVANCE_TIME(20000000); loop();
    ADVANCE_TIME(20000000); loop();
    ADVANCE_TIME(20000000); loop();
    ADVANCE_TIME(20000000); loop();
    ADVANCE_TIME(20000000); loop();
    ADVANCE_TIME(20000000); loop();
    ADVANCE_TIME(20000000); loop();
    ADVANCE_TIME(20000000); loop();
    ADVANCE_TIME(20000000); loop();
    ADVANCE_TIME(20000000); loop();
    ADVANCE_TIME(20000000); loop();
    ADVANCE_TIME(20000000); loop();
    ADVANCE_TIME(20000000); loop();
    ADVANCE_TIME(20000000); loop();
    ADVANCE_TIME(20000000); loop();
    ADVANCE_TIME(20000000); loop();
    ADVANCE_TIME(20000000); loop();
    ADVANCE_TIME(20000000); loop();
    ADVANCE_TIME(20000000); loop();
    ADVANCE_TIME(20000000); loop();
    ADVANCE_TIME(20000000); loop();
    ADVANCE_TIME(20000000); loop();
    ADVANCE_TIME(20000000); loop();
    ADVANCE_TIME(20000000); loop();
    ADVANCE_TIME(20000000); loop();
    ADVANCE_TIME(20000000); loop();
    ADVANCE_TIME(20000000); loop();
    ADVANCE_TIME(20000000); loop();
    ADVANCE_TIME(20000000); loop();
    ADVANCE_TIME(20000000); loop();
    ADVANCE_TIME(20000000); loop();
    ADVANCE_TIME(20000000); loop();
    ADVANCE_TIME(20000000); loop();
    ADVANCE_TIME(20000000); loop();
    ADVANCE_TIME(20000000); loop();
    ADVANCE_TIME(20000000); loop();
    ADVANCE_TIME(20000000); loop();
    ADVANCE_TIME(20000000); loop();
    ADVANCE_TIME(20000000); loop();
    ADVANCE_TIME(20000000); loop();
    ADVANCE_TIME(20000000); loop();
    ADVANCE_TIME(20000000); loop();
    ADVANCE_TIME(20000000); loop();
    ADVANCE_TIME(20000000); loop();
    ADVANCE_TIME(20000000); loop();
    ADVANCE_TIME(20000000); loop();
    ADVANCE_TIME(20000000); loop();
    ADVANCE_TIME(20000000); loop();
    ADVANCE_TIME(20000000); loop();
    ADVANCE_TIME(20000000); loop();
    ADVANCE_TIME(20000000); loop();
    ADVANCE_TIME(20000000); loop();
    ADVANCE_TIME(20000000); loop();
    ADVANCE_TIME(20000000); loop();
    ADVANCE_TIME(20000000); loop();
    ADVANCE_TIME(20000000); loop();
    ADVANCE_TIME(20000000); loop();
    ADVANCE_TIME(20000000); loop();
    ADVANCE_TIME(20000000); loop();
    ADVANCE_TIME(20000000); loop();
    ADVANCE_TIME(20000000); loop();
    ADVANCE_TIME(20000000); loop();
    ADVANCE_TIME(20000000); loop();
    ADVANCE_TIME(20000000); loop();
    ADVANCE_TIME(20000000); loop();
    ADVANCE_TIME(20000000); loop();
    ADVANCE_TIME(20000000); loop();
    ADVANCE_TIME(20000000); loop();
    ADVANCE_TIME(20000000); loop();
    ADVANCE_TIME(20000000); loop();
    ADVANCE_TIME(20000000); loop();
    ADVANCE_TIME(20000000); loop();
    ADVANCE_TIME(20000000); loop();
    ADVANCE_TIME(20000000); loop();
    ADVANCE_TIME(20000000); loop();
    ADVANCE_TIME(20000000); loop();
    ADVANCE_TIME(20000000); loop();
    ADVANCE_TIME(20000000); loop();
    ADVANCE_TIME(20000000); loop();
    ADVANCE_TIME(20000000); loop();
    ADVANCE_TIME(20000000); loop();
    ADVANCE_TIME(20000000); loop();
    ADVANCE_TIME(20000000); loop();
    ADVANCE_TIME(20000000); loop();
    ADVANCE_TIME(20000000); loop();
    ADVANCE_TIME(20000000); loop();
    ADVANCE_TIME(20000000); loop();
    ADVANCE_TIME(20000000); loop();
    ADVANCE_TIME(20000000); loop();
    ADVANCE_TIME(20000000); loop();
    ADVANCE_TIME(20000000); loop();
    ADVANCE_TIME(20000000); loop();
    ADVANCE_TIME(20000000); loop();
    ADVANCE_TIME(20000000); loop();
    ADVANCE_TIME(20000000); loop();
    ADVANCE_TIME(20000000); loop();
    ADVANCE_TIME(20000000); loop();
    ADVANCE_TIME(20000000); loop();
    ADVANCE_TIME(20000000); loop();
    ADVANCE_TIME(20000000); loop();
    ADVANCE_TIME(20000000); loop();
    ADVANCE_TIME(20000000); loop();
    ADVANCE_TIME(20000000); loop();
    ADVANCE_TIME(20000000); loop();
    ADVANCE_TIME(20000000); loop();
    ADVANCE_TIME(20000000); loop();
    ADVANCE_TIME(20000000); loop();
    ADVANCE_TIME(20000000); loop();
    ADVANCE_TIME(20000000); loop();
    ADVANCE_TIME(20000000); loop();
    ADVANCE_TIME(20000000); loop();
    ADVANCE_TIME(20000000); loop();
    ADVANCE_TIME(20000000); loop();
    ADVANCE_TIME(20000000); loop();
    ADVANCE_TIME(20000000); loop();
    ADVANCE_TIME(20000000); loop();
    ADVANCE_TIME(20000000); loop();
    ADVANCE_TIME(20000000); loop();
    ADVANCE_TIME(20000000); loop();
    ADVANCE_TIME(20000000); loop();
    ADVANCE_TIME(20000000); loop();
    ADVANCE_TIME(20000000); loop();
    ADVANCE_TIME(20000000); loop();
    ADVANCE_TIME(20000000); loop();
    ADVANCE_TIME(20000000); loop();
    ADVANCE_TIME(20000000); loop();
    ADVANCE_TIME(20000000); loop();
    ADVANCE_TIME(20000000); loop();
    ADVANCE_TIME(20000000); loop();
    ADVANCE_TIME(20000000); loop();
    ADVANCE_TIME(20000000); loop();
    ADVANCE_TIME(20000000); loop();
    ADVANCE_TIME(20000000); loop();
    ADVANCE_TIME(20000000); loop();
    ADVANCE_TIME(20000000); loop();
    ADVANCE_TIME(20000000); loop();
    ADVANCE_TIME(20000000); loop();
    ADVANCE_TIME(20000000); loop();
    ADVANCE_TIME(20000000); loop();
    ADVANCE_TIME(20000000); loop();
    ADVANCE_TIME(20000000); loop();
    ADVANCE_TIME(20000000); loop();
    ADVANCE_TIME(20000000); loop();
    ADVANCE_TIME(20000000); loop();
    ADVANCE_TIME(20000000); loop();
    ADVANCE_TIME(20000000); loop();
    ADVANCE_TIME(20000000); loop();
    ADVANCE_TIME(20000000); loop();
    ADVANCE_TIME(20000000); loop();
    ADVANCE_TIME(20000000); loop();
    ADVANCE_TIME(20000000); loop();
    ADVANCE_TIME(20000000); loop();
    ADVANCE_TIME(20000000); loop();
    ADVANCE_TIME(20000000); loop();
    ADVANCE_TIME(20000000); loop();
    ADVANCE_TIME(20000000); loop();
    ADVANCE_TIME(20000000); loop();
    ADVANCE_TIME(20000000); loop();
    ADVANCE_TIME(20000000); loop();
    ADVANCE_TIME(20000000); loop();
    ADVANCE_TIME(20000000); loop();
    ADVANCE_TIME(20000000); loop();
    ADVANCE_TIME(20000000); loop();
    ADVANCE_TIME(20000000); loop();
    ADVANCE_TIME(20000000); loop();
    ADVANCE_TIME(20000000); loop();
    ADVANCE_TIME(20000000); loop();
    ADVANCE_TIME(20000000); loop();
    ADVANCE_TIME(20000000); loop();
    ADVANCE_TIME(20000000); loop();
    ADVANCE_TIME(20000000); loop();
    ADVANCE_TIME(20000000); loop();
    ADVANCE_TIME(20000000); loop();
    ADVANCE_TIME(20000000); loop();
    ADVANCE_TIME(20000000); loop();
    ADVANCE_TIME(20000000); loop();
    ADVANCE_TIME(20000000); loop();
    ADVANCE_TIME(20000000); loop();
    ADVANCE_TIME(20000000); loop();
    ADVANCE_TIME(20000000); loop();
    ADVANCE_TIME(20000000); loop();
    ADVANCE_TIME(20000000); loop();
    ADVANCE_TIME(20000000); loop();
    ADVANCE_TIME(20000000); loop();
    ADVANCE_TIME(20000000); loop();
    ADVANCE_TIME(20000000); loop();
    ADVANCE_TIME(20000000); loop();
    ADVANCE_TIME(20000000); loop();
    ADVANCE_TIME(20000000); loop();
    ADVANCE_TIME(20000000); loop();
    ADVANCE_TIME(20000000); loop();
    ADVANCE_TIME(20000000); loop();
    ADVANCE_TIME(20000000); loop();
    ADVANCE_TIME(20000000); loop();
    ADVANCE_TIME(20000000); loop();
    ADVANCE_TIME(20000000); loop();
    ADVANCE_TIME(20000000); loop();
    ADVANCE_TIME(20000000); loop();
    ADVANCE_TIME(20000000); loop();
    ADVANCE_TIME(20000000); loop();
    ADVANCE_TIME(20000000); loop();
    ADVANCE_TIME(20000000); loop();
    ADVANCE_TIME(20000000); loop();
    ADVANCE_TIME(20000000); loop();
    ADVANCE_TIME(20000000); loop();
    ADVANCE_TIME(20000000); loop();
    ADVANCE_TIME(20000000); loop();
    ADVANCE_TIME(20000000); loop();
    ADVANCE_TIME(20000000); loop();
    ADVANCE_TIME(20000000); loop();
    ADVANCE_TIME(20000000); loop();
    ADVANCE_TIME(20000000); loop();
    ADVANCE_TIME(20000000); loop();
    ADVANCE_TIME(20000000); loop();
    ADVANCE_TIME(20000000); loop();
    ADVANCE_TIME(20000000); loop();
    ADVANCE_TIME(20000000); loop();
    ADVANCE_TIME(20000000); loop();
    ADVANCE_TIME(20000000); loop();
    ADVANCE_TIME(20000000); loop();
    ADVANCE_TIME(20000000); loop();
    ADVANCE_TIME(20000000); loop();
    ADVANCE_TIME(20000000); loop();
    ADVANCE_TIME(20000000); loop();
    ADVANCE_TIME(20000000); loop();
    ADVANCE_TIME(20000000); loop();
    ADVANCE_TIME(20000000); loop();
    ADVANCE_TIME(20000000); loop();
    ADVANCE_TIME(20000000); loop();
    ADVANCE_TIME(20000000); loop();
    ADVANCE_TIME(20000000); loop();
    ADVANCE_TIME(20000000); loop();
    ADVANCE_TIME(20000000); loop();
    ADVANCE_TIME(20000000); loop();
    ADVANCE_TIME(20000000); loop();
    ADVANCE_TIME(20000000); loop();
    ADVANCE_TIME(20000000); loop();
    ADVANCE_TIME(20000000); loop();
    ADVANCE_TIME(20000000); loop();
    ADVANCE_TIME(20000000); loop();
    ADVANCE_TIME(20000000); loop();
    ADVANCE_TIME(20000000); loop();
    ADVANCE_TIME(20000000); loop();
    ADVANCE_TIME(20000000); loop();
    ADVANCE_TIME(20000000); loop();
    ADVANCE_TIME(20000000); loop();
    ADVANCE_TIME(20000000); loop();
    ADVANCE_TIME(20000000); loop();
    ADVANCE_TIME(20000000); loop();
    ADVANCE_TIME(20000000); loop();
    ADVANCE_TIME(20000000); loop();
    ADVANCE_TIME(20000000); loop();
    ADVANCE_TIME(20000000); loop();
    ADVANCE_TIME(20000000); loop();
    ADVANCE_TIME(20000000); loop();
    ADVANCE_TIME(20000000); loop();
    ADVANCE_TIME(20000000); loop();
    ADVANCE_TIME(20000000); loop();
    ADVANCE_TIME(20000000); loop();
    ADVANCE_TIME(20000000); loop();
    ADVANCE_TIME(20000000); loop();
    ADVANCE_TIME(20000000); loop();
    ADVANCE_TIME(20000000); loop();
    ADVANCE_TIME(20000000); loop();
    ADVANCE_TIME(20000000); loop();
    ADVANCE_TIME(20000000); loop();
    ADVANCE_TIME(20000000); loop();
    ADVANCE_TIME(20000000); loop();
    ADVANCE_TIME(20000000); loop();
    ADVANCE_TIME(20000000); loop();
    ADVANCE_TIME(20000000); loop();
    ADVANCE_TIME(20000000); loop();
    ADVANCE_TIME(20000000); loop();
    ADVANCE_TIME(20000000); loop();
    ADVANCE_TIME(20000000); loop();
    ADVANCE_TIME(20000000); loop();
    ADVANCE_TIME(20000000); loop();
    ADVANCE_TIME(20000000); loop();
    ADVANCE_TIME(20000000); loop();
    ADVANCE_TIME(20000000); loop();
    ADVANCE_TIME(20000000); loop();
    ADVANCE_TIME(20000000); loop();
    ADVANCE_TIME(20000000); loop();
    ADVANCE_TIME(20000000); loop();
    ADVANCE_TIME(20000000); loop();
    ADVANCE_TIME(20000000); loop();
    ADVANCE_TIME(20000000); loop();
    ADVANCE_TIME(20000000); loop();
    ADVANCE_TIME(20000000); loop();
    ADVANCE_TIME(20000000); loop();
    ADVANCE_TIME(20000000); loop();
    ADVANCE_TIME(20000000); loop();
    ADVANCE_TIME(20000000); loop();
    ADVANCE_TIME(20000000); loop();
    ADVANCE_TIME(20000000); loop();
    ADVANCE_TIME(20000000); loop();
    ADVANCE_TIME(20000000); loop();
    ADVANCE_TIME(20000000); loop();
    ADVANCE_TIME(20000000); loop();
    ADVANCE_TIME(20000000); loop();
    ADVANCE_TIME(20000000); loop();
    ADVANCE_TIME(20000000); loop();
    ADVANCE_TIME(20000000); loop();
    ADVANCE_TIME(20000000); loop();
    ADVANCE_TIME(20000000); loop();
    ADVANCE_TIME(20000000); loop();
    ADVANCE_TIME(20000000); loop();
    ADVANCE_TIME(20000000); loop();
    ADVANCE_TIME(20000000); loop();
    ADVANCE_TIME(20000000); loop();
    ADVANCE_TIME(20000000); loop();
    ADVANCE_TIME(20000000); loop();
    ADVANCE_TIME(20000000); loop();
    ADVANCE_TIME(20000000); loop();
    ADVANCE_TIME(20000000); loop();
    ADVANCE_TIME(20000000); loop();
    ADVANCE_TIME(20000000); loop();
    ADVANCE_TIME(20000000); loop();
    ADVANCE_TIME(20000000); loop();
    ADVANCE_TIME(20000000); loop();
    ADVANCE_TIME(20000000); loop();
    ADVANCE_TIME(20000000); loop();
    ADVANCE_TIME(20000000); loop();
    ADVANCE_TIME(20000000); loop();
    ADVANCE_TIME(20000000); loop();
    ADVANCE_TIME(20000000); loop();
    ADVANCE_TIME(20000000); loop();
    ADVANCE_TIME(20000000); loop();
    ADVANCE_TIME(20000000); loop();
    ADVANCE_TIME(20000000); loop();
    ADVANCE_TIME(20000000); loop();
    ADVANCE_TIME(20000000); loop();
    ADVANCE_TIME(20000000); loop();
    ADVANCE_TIME(20000000); loop();
    ADVANCE_TIME(20000000); loop();
    ADVANCE_TIME(20000000); loop();
    ADVANCE_TIME(20000000); loop();
    ADVANCE_TIME(20000000); loop();
    ADVANCE_TIME(20000000); loop();
    ADVANCE_TIME(20000000); loop();
    ADVANCE_TIME(20000000); loop();
    ADVANCE_TIME(20000000); loop();
    ADVANCE_TIME(20000000); loop();
    ADVANCE_TIME(20000000); loop();
    ADVANCE_TIME(20000000); loop();
    ADVANCE_TIME(20000000); loop();
    ADVANCE_TIME(20000000); loop();
    ADVANCE_TIME(20000000); loop();
    ADVANCE_TIME(20000000); loop();
    ADVANCE_TIME(20000000); loop();
    ADVANCE_TIME(20000000); loop();
    ADVANCE_TIME(20000000); loop();
    ADVANCE_TIME(20000000); loop();
    ADVANCE_TIME(20000000); loop();
    ADVANCE_TIME(20000000); loop();
    ADVANCE_TIME(20000000); loop();
    ADVANCE_TIME(20000000); loop();
    ADVANCE_TIME(20000000); loop();
    ADVANCE_TIME(20000000); loop();
    ADVANCE_TIME(20000000); loop();
    ADVANCE_TIME(20000000); loop();
    ADVANCE_TIME(20000000); loop();
    ADVANCE_TIME(20000000); loop();
    ADVANCE_TIME(20000000); loop();
    ADVANCE_TIME(20000000); loop();
    ADVANCE_TIME(20000000); loop();
    ADVANCE_TIME(20000000); loop();
    ADVANCE_TIME(20000000); loop();
    ADVANCE_TIME(20000000); loop();
    ADVANCE_TIME(20000000); loop();
    ADVANCE_TIME(20000000); loop();
    ADVANCE_TIME(20000000); loop();
    ADVANCE_TIME(20000000); loop();
    ADVANCE_TIME(20000000); loop();
    ADVANCE_TIME(20000000); loop();
    ADVANCE_TIME(20000000); loop();
    ADVANCE_TIME(20000000); loop();
    ADVANCE_TIME(20000000); loop();
    ADVANCE_TIME(20000000); loop();
    ADVANCE_TIME(20000000); loop();
    ADVANCE_TIME(20000000); loop();
    ADVANCE_TIME(20000000); loop();
    ADVANCE_TIME(20000000); loop();
    ADVANCE_TIME(20000000); loop();
    ADVANCE_TIME(20000000); loop();
    ADVANCE_TIME(20000000); loop();
    ADVANCE_TIME(20000000); loop();
    ADVANCE_TIME(20000000); loop();
    ADVANCE_TIME(20000000); loop();
    ADVANCE_TIME(20000000); loop();
    ADVANCE_TIME(20000000); loop();
    ADVANCE_TIME(20000000); loop();
    ADVANCE_TIME(20000000); loop();
    ADVANCE_TIME(20000000); loop();
    ADVANCE_TIME(20000000); loop();
    ADVANCE_TIME(20000000); loop();
    ADVANCE_TIME(20000000); loop();
    ADVANCE_TIME(20000000); loop();
    ADVANCE_TIME(20000000); loop();
    ADVANCE_TIME(20000000); loop();
    ADVANCE_TIME(20000000); loop();
    ADVANCE_TIME(20000000); loop();
    ADVANCE_TIME(20000000); loop();
    ADVANCE_TIME(20000000); loop();
    ADVANCE_TIME(20000000); loop();
    ADVANCE_TIME(20000000); loop();
    ADVANCE_TIME(20000000); loop();
    ADVANCE_TIME(20000000); loop();
    ADVANCE_TIME(20000000); loop();
    ADVANCE_TIME(20000000); loop();
    ADVANCE_TIME(20000000); loop();
    ADVANCE_TIME(20000000); loop();
    ADVANCE_TIME(20000000); loop();
    ADVANCE_TIME(20000000); loop();
    ADVANCE_TIME(20000000); loop();
    ADVANCE_TIME(20000000); loop();
    ADVANCE_TIME(20000000); loop();
    ADVANCE_TIME(20000000); loop();
    ADVANCE_TIME(20000000); loop();
    ADVANCE_TIME(20000000); loop();
    ADVANCE_TIME(20000000); loop();
    ADVANCE_TIME(20000000); loop();
    ADVANCE_TIME(20000000); loop();
    ADVANCE_TIME(20000000); loop();
    ADVANCE_TIME(20000000); loop();
    ADVANCE_TIME(20000000); loop();
    ADVANCE_TIME(20000000); loop();
    ADVANCE_TIME(20000000); loop();
    ADVANCE_TIME(20000000); loop();
    ADVANCE_TIME(20000000); loop();
    ADVANCE_TIME(20000000); loop();
    ADVANCE_TIME(20000000); loop();
    ADVANCE_TIME(20000000); loop();
    ADVANCE_TIME(20000000); loop();
    ADVANCE_TIME(20000000); loop();
    ADVANCE_TIME(20000000); loop();
    ADVANCE_TIME(20000000); loop();
    ADVANCE_TIME(20000000); loop();
    ADVANCE_TIME(20000000); loop();
    ADVANCE_TIME(20000000); loop();
    ADVANCE_TIME(20000000); loop();
    ADVANCE_TIME(20000000); loop();
    ADVANCE_TIME(20000000); loop();
    ADVANCE_TIME(20000000); loop();
    ADVANCE_TIME(20000000); loop();
    ADVANCE_TIME(20000000); loop();
    ADVANCE_TIME(20000000); loop();
    ADVANCE_TIME(20000000); loop();
    ADVANCE_TIME(20000000); loop();
    ADVANCE_TIME(20000000); loop();
    ADVANCE_TIME(20000000); loop();
    ADVANCE_TIME(20000000); loop();
    ADVANCE_TIME(20000000); loop();
    ADVANCE_TIME(20000000); loop();
    ADVANCE_TIME(20000000); loop();
    ADVANCE_TIME(20000000); loop();
    ADVANCE_TIME(20000000); loop();
    ADVANCE_TIME(20000000); loop();
    ADVANCE_TIME(20000000); loop();
    ADVANCE_TIME(20000000); loop();
    ADVANCE_TIME(20000000); loop();
    ADVANCE_TIME(20000000); loop();
    ADVANCE_TIME(20000000); loop();
    ADVANCE_TIME(20000000); loop();
    ADVANCE_TIME(20000000); loop();
    ADVANCE_TIME(20000000); loop();
    ADVANCE_TIME(20000000); loop();
    ADVANCE_TIME(20000000); loop();
    ADVANCE_TIME(20000000); loop();
    ADVANCE_TIME(20000000); loop();
    ADVANCE_TIME(20000000); loop();
    ADVANCE_TIME(20000000); loop();
    ADVANCE_TIME(20000000); loop();
    ADVANCE_TIME(20000000); loop();
    ADVANCE_TIME(20000000); loop();
    ADVANCE_TIME(20000000); loop();
    ADVANCE_TIME(20000000); loop();
    ADVANCE_TIME(20000000); loop();
    ADVANCE_TIME(20000000); loop();
    ADVANCE_TIME(20000000); loop();
    ADVANCE_TIME(20000000); loop();
    ADVANCE_TIME(20000000); loop();
    ADVANCE_TIME(20000000); loop();
    ADVANCE_TIME(20000000); loop();
    ADVANCE_TIME(20000000); loop();
    ADVANCE_TIME(20000000); loop();
    ADVANCE_TIME(20000000); loop();
    ADVANCE_TIME(20000000); loop();
    ADVANCE_TIME(20000000); loop();
    ADVANCE_TIME(20000000); loop();
    ADVANCE_TIME(20000000); loop();
    ADVANCE_TIME(20000000); loop();
    ADVANCE_TIME(20000000); loop();
    ADVANCE_TIME(20000000); loop();
    ADVANCE_TIME(20000000); loop();
    ADVANCE_TIME(20000000); loop();
    ADVANCE_TIME(20000000); loop();
    ADVANCE_TIME(20000000); loop();
    ADVANCE_TIME(20000000); loop();
    ADVANCE_TIME(20000000); loop();
    ADVANCE_TIME(20000000); loop();
    ADVANCE_TIME(20000000); loop();
    ADVANCE_TIME(20000000); loop();
    ADVANCE_TIME(20000000); loop();
    ADVANCE_TIME(20000000); loop();
    ADVANCE_TIME(20000000); loop();
    ADVANCE_TIME(20000000); loop();
    ADVANCE_TIME(20000000); loop();
    ADVANCE_TIME(20000000); loop();
    ADVANCE_TIME(20000000); loop();
    ADVANCE_TIME(20000000); loop();
    ADVANCE_TIME(20000000); loop();
    ADVANCE_TIME(20000000); loop();
    ADVANCE_TIME(20000000); loop();
    ADVANCE_TIME(20000000); loop();
    ADVANCE_TIME(20000000); loop();
    ADVANCE_TIME(20000000); loop();
    ADVANCE_TIME(20000000); loop();
    ADVANCE_TIME(20000000); loop();
    ADVANCE_TIME(20000000); loop();
    ADVANCE_TIME(20000000); loop();
    ADVANCE_TIME(20000000); loop();
    ADVANCE_TIME(20000000); loop();
    ADVANCE_TIME(20000000); loop();
    ADVANCE_TIME(20000000); loop();
    ADVANCE_TIME(20000000); loop();
    ADVANCE_TIME(20000000); loop();
    ADVANCE_TIME(20000000); loop();
    ADVANCE_TIME(20000000); loop();
    ADVANCE_TIME(20000000); loop();
    ADVANCE_TIME(20000000); loop();
    ADVANCE_TIME(20000000); loop();
    ADVANCE_TIME(20000000); loop();
    ADVANCE_TIME(20000000); loop();
    ADVANCE_TIME(20000000); loop();
    ADVANCE_TIME(20000000); loop();
    ADVANCE_TIME(20000000); loop();
    ADVANCE_TIME(20000000); loop();
    ADVANCE_TIME(20000000); loop();
    ADVANCE_TIME(20000000); loop();
    ADVANCE_TIME(20000000); loop();
    ADVANCE_TIME(20000000); loop();
    ADVANCE_TIME(20000000); loop();
    ADVANCE_TIME(20000000); loop();
    ADVANCE_TIME(20000000); loop();
    ADVANCE_TIME(20000000); loop();
    ADVANCE_TIME(20000000); loop();
    ADVANCE_TIME(20000000); loop();
    ADVANCE_TIME(20000000); loop();
    ADVANCE_TIME(20000000); loop();
    ADVANCE_TIME(20000000); loop();
    ADVANCE_TIME(20000000); loop();
    ADVANCE_TIME(20000000); loop();
    ADVANCE_TIME(20000000); loop();
    ADVANCE_TIME(20000000); loop();
    ADVANCE_TIME(20000000); loop();
    ADVANCE_TIME(20000000); loop();
    ADVANCE_TIME(20000000); loop();
    ADVANCE_TIME(20000000); loop();
    ADVANCE_TIME(20000000); loop();
    ADVANCE_TIME(20000000); loop();
    ADVANCE_TIME(20000000); loop();
    ADVANCE_TIME(20000000); loop();
    ADVANCE_TIME(20000000); loop();
    ADVANCE_TIME(20000000); loop();
    ADVANCE_TIME(20000000); loop();
    ADVANCE_TIME(20000000); loop();
    ADVANCE_TIME(20000000); loop();
    ADVANCE_TIME(20000000); loop();
    ADVANCE_TIME(20000000); loop();
    ADVANCE_TIME(20000000); loop();
    ADVANCE_TIME(20000000); loop();
    ADVANCE_TIME(20000000); loop();
    ADVANCE_TIME(20000000); loop();
    ADVANCE_TIME(20000000); loop();
    ADVANCE_TIME(20000000); loop();
    ADVANCE_TIME(20000000); loop();
    ADVANCE_TIME(20000000); loop();
    ADVANCE_TIME(20000000); loop();
    ADVANCE_TIME(20000000); loop();
    ADVANCE_TIME(20000000); loop();
    ADVANCE_TIME(20000000); loop();
    ADVANCE_TIME(20000000); loop();
    ADVANCE_TIME(20000000); loop();
    ADVANCE_TIME(20000000); loop();
    ADVANCE_TIME(20000000); loop();
    ADVANCE_TIME(20000000); loop();
    ADVANCE_TIME(20000000); loop();
    ADVANCE_TIME(20000000); loop();
    ADVANCE_TIME(20000000); loop();
    ADVANCE_TIME(20000000); loop();
    ADVANCE_TIME(20000000); loop();
    ADVANCE_TIME(20000000); loop();
    ADVANCE_TIME(20000000); loop();
    ADVANCE_TIME(20000000); loop();
    ADVANCE_TIME(20000000); loop();
    ADVANCE_TIME(20000000); loop();
    ADVANCE_TIME(20000000); loop();
    ADVANCE_TIME(20000000); loop();
    ADVANCE_TIME(20000000); loop();
    ADVANCE_TIME(20000000); loop();
    ADVANCE_TIME(20000000); loop();
    ADVANCE_TIME(20000000); loop();
    ADVANCE_TIME(20000000); loop();
    ADVANCE_TIME(20000000); loop();
    ADVANCE_TIME(20000000); loop();
    ADVANCE_TIME(20000000); loop();
    ADVANCE_TIME(20000000); loop();
    ADVANCE_TIME(20000000); loop();
    ADVANCE_TIME(20000000); loop();
    ADVANCE_TIME(20000000); loop();
    ADVANCE_TIME(20000000); loop();
    ADVANCE_TIME(20000000); loop();
    ADVANCE_TIME(20000000); loop();
    ADVANCE_TIME(20000000); loop();
    ADVANCE_TIME(20000000); loop();
    ADVANCE_TIME(20000000); loop();
    ADVANCE_TIME(20000000); loop();
    ADVANCE_TIME(20000000); loop();
    ADVANCE_TIME(20000000); loop();
    ADVANCE_TIME(20000000); loop();
    ADVANCE_TIME(20000000); loop();
    ADVANCE_TIME(20000000); loop();
    ADVANCE_TIME(20000000); loop();
    ADVANCE_TIME(20000000); loop();
    ADVANCE_TIME(20000000); loop();
    ADVANCE_TIME(20000000); loop();
    ADVANCE_TIME(20000000); loop();
    ADVANCE_TIME(20000000); loop();
    ADVANCE_TIME(20000000); loop();
    ADVANCE_TIME(20000000); loop();
    ADVANCE_TIME(20000000); loop();
    ADVANCE_TIME(20000000); loop();
    ADVANCE_TIME(20000000); loop();
    ADVANCE_TIME(20000000); loop();
    ADVANCE_TIME(20000000); loop();
    ADVANCE_TIME(20000000); loop();
    ADVANCE_TIME(20000000); loop();
    ADVANCE_TIME(20000000); loop();
    ADVANCE_TIME(20000000); loop();
    ADVANCE_TIME(20000000); loop();
    ADVANCE_TIME(20000000); loop();
    ADVANCE_TIME(20000000); loop();
    ADVANCE_TIME(20000000); loop();
    ADVANCE_TIME(20000000); loop();
    ADVANCE_TIME(20000000); loop();
    ADVANCE_TIME(20000000); loop();
    ADVANCE_TIME(20000000); loop();
    ADVANCE_TIME(20000000); loop();
    ADVANCE_TIME(20000000); loop();
    ADVANCE_TIME(20000000); loop();
    ADVANCE_TIME(20000000); loop();
    ADVANCE_TIME(20000000); loop();
    ADVANCE_TIME(20000000); loop();
    ADVANCE_TIME(20000000); loop();
    ADVANCE_TIME(20000000); loop();
    ADVANCE_TIME(20000000); loop();
    ADVANCE_TIME(20000000); loop();
    ADVANCE_TIME(20000000); loop();
    ADVANCE_TIME(20000000); loop();
    ADVANCE_TIME(20000000); loop();
    ADVANCE_TIME(20000000); loop();
    ADVANCE_TIME(20000000); loop();
    ADVANCE_TIME(20000000); loop();
    ADVANCE_TIME(20000000); loop();
    ADVANCE_TIME(20000000); loop();
    ADVANCE_TIME(20000000); loop();
    ADVANCE_TIME(20000000); loop();
    ADVANCE_TIME(20000000); loop();
    ADVANCE_TIME(20000000); loop();
    ADVANCE_TIME(20000000); loop();
    ADVANCE_TIME(20000000); loop();
    ADVANCE_TIME(20000000); loop();
    ADVANCE_TIME(20000000); loop();
    ADVANCE_TIME(20000000); loop();
    ADVANCE_TIME(20000000); loop();
    ADVANCE_TIME(20000000); loop();
    ADVANCE_TIME(20000000); loop();
    ADVANCE_TIME(20000000); loop();
    ADVANCE_TIME(20000000); loop();
    ADVANCE_TIME(20000000); loop();
    ADVANCE_TIME(20000000); loop();
    ADVANCE_TIME(20000000); loop();
    ADVANCE_TIME(20000000); loop();
    ADVANCE_TIME(20000000); loop();
    ADVANCE_TIME(20000000); loop();
    ADVANCE_TIME(20000000); loop();
    ADVANCE_TIME(20000000); loop();
    ADVANCE_TIME(20000000); loop();
    ADVANCE_TIME(20000000); loop();
    ADVANCE_TIME(20000000); loop();
    ADVANCE_TIME(20000000); loop();
    ADVANCE_TIME(20000000); loop();
    ADVANCE_TIME(20000000); loop();
    ADVANCE_TIME(20000000); loop();
    ADVANCE_TIME(20000000); loop();
    ADVANCE_TIME(20000000); loop();
    ADVANCE_TIME(20000000); loop();
    ADVANCE_TIME(20000000); loop();
    ADVANCE_TIME(20000000); loop();
    ADVANCE_TIME(20000000); loop();
    ADVANCE_TIME(20000000); loop();
    ADVANCE_TIME(20000000); loop();
    ADVANCE_TIME(20000000); loop();
    ADVANCE_TIME(20000000); loop();
    ADVANCE_TIME(20000000); loop();
    ADVANCE_TIME(20000000); loop();
    ADVANCE_TIME(20000000); loop();
    ADVANCE_TIME(20000000); loop();
    ADVANCE_TIME(20000000); loop();
    ADVANCE_TIME(20000000); loop();
    ADVANCE_TIME(20000000); loop();
    ADVANCE_TIME(20000000); loop();
    ADVANCE_TIME(20000000); loop();
    ADVANCE_TIME(20000000); loop();
    ADVANCE_TIME(20000000); loop();
    ADVANCE_TIME(20000000); loop();
    ADVANCE_TIME(20000000); loop();
    ADVANCE_TIME(20000000); loop();
    ADVANCE_TIME(20000000); loop();
    ADVANCE_TIME(20000000); loop();
    ADVANCE_TIME(20000000); loop();
    ADVANCE_TIME(20000000); loop();
    ADVANCE_TIME(20000000); loop();
    ADVANCE_TIME(20000000); loop();
    ADVANCE_TIME(20000000); loop();
    ADVANCE_TIME(20000000); loop();
    ADVANCE_TIME(20000000); loop();
    ADVANCE_TIME(20000000); loop();
    ADVANCE_TIME(20000000); loop();
    ADVANCE_TIME(20000000); loop();
    ADVANCE_TIME(20000000); loop();
    ADVANCE_TIME(20000000); loop();
    ADVANCE_TIME(20000000); loop();
    ADVANCE_TIME(20000000); loop();
    ADVANCE_TIME(20000000); loop();
    ADVANCE_TIME(20000000); loop();
    ADVANCE_TIME(20000000); loop();
    ADVANCE_TIME(20000000); loop();
    ADVANCE_TIME(20000000); loop();
    ADVANCE_TIME(20000000); loop();
    ADVANCE_TIME(20000000); loop();
    ADVANCE_TIME(20000000); loop();
    ADVANCE_TIME(20000000); loop();
    ADVANCE_TIME(20000000); loop();
    ADVANCE_TIME(20000000); loop();
    ADVANCE_TIME(20000000); loop();
    ADVANCE_TIME(20000000); loop();
    ADVANCE_TIME(20000000); loop();
    ADVANCE_TIME(20000000); loop();
    ADVANCE_TIME(20000000); loop();
    ADVANCE_TIME(20000000); loop();
    ADVANCE_TIME(20000000); loop();
    ADVANCE_TIME(20000000); loop();
    ADVANCE_TIME(20000000); loop();
    ADVANCE_TIME(20000000); loop();
    ADVANCE_TIME(20000000); loop();
    ADVANCE_TIME(20000000); loop();
    ADVANCE_TIME(20000000); loop();
    ADVANCE_TIME(20000000); loop();
    ADVANCE_TIME(20000000); loop();
    ADVANCE_TIME(20000000); loop();
    ADVANCE_TIME(20000000); loop();
    ADVANCE_TIME(20000000); loop();
    ADVANCE_TIME(20000000); loop();
    ADVANCE_TIME(20000000); loop();
    ADVANCE_TIME(20000000); loop();
    ADVANCE_TIME(20000000); loop();
    ADVANCE_TIME(20000000); loop();
    ADVANCE_TIME(20000000); loop();
    ADVANCE_TIME(20000000); loop();
    ADVANCE_TIME(20000000); loop();
    ADVANCE_TIME(20000000); loop();
    ADVANCE_TIME(20000000); loop();
    ADVANCE_TIME(20000000); loop();
    ADVANCE_TIME(20000000); loop();
    ADVANCE_TIME(20000000); loop();
    ADVANCE_TIME(20000000); loop();
    ADVANCE_TIME(20000000); loop();
    ADVANCE_TIME(20000000); loop();
    ADVANCE_TIME(20000000); loop();
    ADVANCE_TIME(20000000); loop();
    ADVANCE_TIME(20000000); loop();
    ADVANCE_TIME(20000000); loop();
    ADVANCE_TIME(20000000); loop();
    ADVANCE_TIME(20000000); loop();
    ADVANCE_TIME(20000000); loop();
    ADVANCE_TIME(20000000); loop();
    ADVANCE_TIME(20000000); loop();
    ADVANCE_TIME(20000000); loop();
    ADVANCE_TIME(20000000); loop();
    ADVANCE_TIME(20000000); loop();
    ADVANCE_TIME(20000000); loop();
    ADVANCE_TIME(20000000); loop();
    ADVANCE_TIME(20000000); loop();
    ADVANCE_TIME(20000000); loop();
    ADVANCE_TIME(20000000); loop();
    ADVANCE_TIME(20000000); loop();
    ADVANCE_TIME(20000000); loop();
    ADVANCE_TIME(20000000); loop();
    ADVANCE_TIME(20000000); loop();
    ADVANCE_TIME(20000000); loop();
    ADVANCE_TIME(20000000); loop();
    ADVANCE_TIME(20000000); loop();
    ADVANCE_TIME(20000000); loop();
    ADVANCE_TIME(20000000); loop();
    ADVANCE_TIME(20000000); loop();
    ADVANCE_TIME(20000000); loop();
    ADVANCE_TIME(20000000); loop();
    ADVANCE_TIME(20000000); loop();
    ADVANCE_TIME(20000000); loop();
    ADVANCE_TIME(20000000); loop();
    ADVANCE_TIME(20000000); loop();
    ADVANCE_TIME(20000000); loop();
    ADVANCE_TIME(20000000); loop();
    ADVANCE_TIME(20000000); loop();
    ADVANCE_TIME(20000000); loop();
    ADVANCE_TIME(20000000); loop();
    ADVANCE_TIME(20000000); loop();
    ADVANCE_TIME(20000000); loop();
    ADVANCE_TIME(20000000); loop();
    ADVANCE_TIME(20000000); loop();
    ADVANCE_TIME(20000000); loop();
    ADVANCE_TIME(20000000); loop();
    ADVANCE_TIME(20000000); loop();
    ADVANCE_TIME(20000000); loop();
    ADVANCE_TIME(20000000); loop();
    ADVANCE_TIME(20000000); loop();
    ADVANCE_TIME(20000000); loop();
    ADVANCE_TIME(20000000); loop();
    ADVANCE_TIME(20000000); loop();
    ADVANCE_TIME(20000000); loop();
    ADVANCE_TIME(20000000); loop();
    ADVANCE_TIME(20000000); loop();
    ADVANCE_TIME(20000000); loop();
    ADVANCE_TIME(20000000); loop();
    ADVANCE_TIME(20000000); loop();
    ADVANCE_TIME(20000000); loop();
    ADVANCE_TIME(20000000); loop();
    ADVANCE_TIME(20000000); loop();
    ADVANCE_TIME(20000000); loop();
    ADVANCE_TIME(20000000); loop();
    ADVANCE_TIME(20000000); loop();
    ADVANCE_TIME(20000000); loop();
    ADVANCE_TIME(20000000); loop();
    ADVANCE_TIME(20000000); loop();
    ADVANCE_TIME(20000000); loop();
    ADVANCE_TIME(20000000); loop();
    ADVANCE_TIME(20000000); loop();
    ADVANCE_TIME(20000000); loop();
    ADVANCE_TIME(20000000); loop();
    ADVANCE_TIME(20000000); loop();
    ADVANCE_TIME(20000000); loop();
    ADVANCE_TIME(20000000); loop();
    ADVANCE_TIME(20000000); loop();
    ADVANCE_TIME(20000000); loop();
    ADVANCE_TIME(20000000); loop();
    ADVANCE_TIME(20000000); loop();
    ADVANCE_TIME(20000000); loop();
    ADVANCE_TIME(20000000); loop();
    ADVANCE_TIME(20000000); loop();
    ADVANCE_TIME(20000000); loop();
    ADVANCE_TIME(20000000); loop();
    ADVANCE_TIME(20000000); loop();
    ADVANCE_TIME(20000000); loop();
    ADVANCE_TIME(20000000); loop();
    ADVANCE_TIME(20000000); loop();
    ADVANCE_TIME(20000000); loop();
    ADVANCE_TIME(20000000); loop();
    ADVANCE_TIME(20000000); loop();
    ADVANCE_TIME(20000000); loop();
    ADVANCE_TIME(20000000); loop();
    ADVANCE_TIME(20000000); loop();
    ADVANCE_TIME(20000000); loop();
    ADVANCE_TIME(20000000); loop();
    ADVANCE_TIME(20000000); loop();
    ADVANCE_TIME(20000000); loop();
    ADVANCE_TIME(20000000); loop();
    ADVANCE_TIME(20000000); loop();
    ADVANCE_TIME(20000000); loop();
    ADVANCE_TIME(20000000); loop();
    ADVANCE_TIME(20000000); loop();
    ADVANCE_TIME(20000000); loop();
    ADVANCE_TIME(20000000); loop();
    ADVANCE_TIME(20000000); loop();
    ADVANCE_TIME(20000000); loop();
    ADVANCE_TIME(20000000); loop();
    ADVANCE_TIME(20000000); loop();
    ADVANCE_TIME(20000000); loop();
    ADVANCE_TIME(20000000); loop();
    ADVANCE_TIME(20000000); loop();
    ADVANCE_TIME(20000000); loop();
    ADVANCE_TIME(20000000); loop();
    ADVANCE_TIME(20000000); loop();
    ADVANCE_TIME(20000000); loop();
    ADVANCE_TIME(20000000); loop();
    ADVANCE_TIME(20000000); loop();
    ADVANCE_TIME(20000000); loop();
    ADVANCE_TIME(20000000); loop();
    ADVANCE_TIME(20000000); loop();
    ADVANCE_TIME(20000000); loop();
    ADVANCE_TIME(20000000); loop();
    ADVANCE_TIME(20000000); loop();
    ADVANCE_TIME(20000000); loop();
    ADVANCE_TIME(20000000); loop();
    ADVANCE_TIME(20000000); loop();
    ADVANCE_TIME(20000000); loop();
    ADVANCE_TIME(20000000); loop();
    ADVANCE_TIME(20000000); loop();
    ADVANCE_TIME(20000000); loop();
    ADVANCE_TIME(20000000); loop();
    ADVANCE_TIME(20000000); loop();
    ADVANCE_TIME(20000000); loop();
    ADVANCE_TIME(20000000); loop();
    ADVANCE_TIME(20000000); loop();
    ADVANCE_TIME(20000000); loop();
    ADVANCE_TIME(20000000); loop();
    ADVANCE_TIME(20000000); loop();
    ADVANCE_TIME(20000000); loop();
    ADVANCE_TIME(20000000); loop();
    ADVANCE_TIME(20000000); loop();
    ADVANCE_TIME(20000000); loop();
    ADVANCE_TIME(20000000); loop();
    ADVANCE_TIME(20000000); loop();
    ADVANCE_TIME(20000000); loop();
    ADVANCE_TIME(20000000); loop();
    ADVANCE_TIME(20000000); loop();
    ADVANCE_TIME(20000000); loop();
    ADVANCE_TIME(20000000); loop();
    ADVANCE_TIME(20000000); loop();
    ADVANCE_TIME(20000000); loop();
    ADVANCE_TIME(20000000); loop();
    ADVANCE_TIME(20000000); loop();
    ADVANCE_TIME(20000000); loop();
    ADVANCE_TIME(20000000); loop();
    ADVANCE_TIME(20000000); loop();
    ADVANCE_TIME(20000000); loop();
    ADVANCE_TIME(20000000); loop();
    ADVANCE_TIME(20000000); loop();
    ADVANCE_TIME(20000000); loop();
    ADVANCE_TIME(20000000); loop();
    ADVANCE_TIME(20000000); loop();
    ADVANCE_TIME(20000000); loop();
    ADVANCE_TIME(20000000); loop();
    ADVANCE_TIME(20000000); loop();
    ADVANCE_TIME(20000000); loop();
    ADVANCE_TIME(20000000); loop();
    ADVANCE_TIME(20000000); loop();
    ADVANCE_TIME(20000000); loop();
    ADVANCE_TIME(20000000); loop();
    ADVANCE_TIME(20000000); loop();
    ADVANCE_TIME(20000000); loop();
    ADVANCE_TIME(20000000); loop();
    ADVANCE_TIME(20000000); loop();
    ADVANCE_TIME(20000000); loop();
    ADVANCE_TIME(20000000); loop();
    ADVANCE_TIME(20000000); loop();
    ADVANCE_TIME(20000000); loop();
    ADVANCE_TIME(20000000); loop();
    ADVANCE_TIME(20000000); loop();
    ADVANCE_TIME(20000000); loop();
    ADVANCE_TIME(20000000); loop();
    ADVANCE_TIME(20000000); loop();
    ADVANCE_TIME(20000000); loop();
    ADVANCE_TIME(20000000); loop();
    ADVANCE_TIME(20000000); loop();
    ADVANCE_TIME(20000000); loop();
    ADVANCE_TIME(20000000); loop();
    ADVANCE_TIME(20000000); loop();
    ADVANCE_TIME(20000000); loop();
    ADVANCE_TIME(20000000); loop();
    ADVANCE_TIME(20000000); loop();
    ADVANCE_TIME(20000000); loop();
    ADVANCE_TIME(20000000); loop();
    ADVANCE_TIME(20000000); loop();
    ADVANCE_TIME(20000000); loop();
    ADVANCE_TIME(20000000); loop();
    ADVANCE_TIME(20000000); loop();
    ADVANCE_TIME(20000000); loop();
    ADVANCE_TIME(20000000); loop();
    ADVANCE_TIME(20000000); loop();
    ADVANCE_TIME(20000000); loop();
    ADVANCE_TIME(20000000); loop();
    ADVANCE_TIME(20000000); loop();
    ADVANCE_TIME(20000000); loop();
    ADVANCE_TIME(20000000); loop();
    ADVANCE_TIME(20000000); loop();
    ADVANCE_TIME(20000000); loop();
    ADVANCE_TIME(20000000); loop();
    ADVANCE_TIME(20000000); loop();
    ADVANCE_TIME(20000000); loop();
    ADVANCE_TIME(20000000); loop();
    ADVANCE_TIME(20000000); loop();
    ADVANCE_TIME(20000000); loop();
    ADVANCE_TIME(20000000); loop();
    ADVANCE_TIME(20000000); loop();
    ADVANCE_TIME(20000000); loop();
    ADVANCE_TIME(20000000); loop();
    ADVANCE_TIME(20000000); loop();
    ADVANCE_TIME(20000000); loop();
    ADVANCE_TIME(20000000); loop();
    ADVANCE_TIME(20000000); loop();
    ADVANCE_TIME(20000000); loop();
    ADVANCE_TIME(20000000); loop();
    ADVANCE_TIME(20000000); loop();
    ADVANCE_TIME(20000000); loop();
    ADVANCE_TIME(20000000); loop();
    ADVANCE_TIME(20000000); loop();
    ADVANCE_TIME(20000000); loop();
    ADVANCE_TIME(20000000); loop();
    ADVANCE_TIME(20000000); loop();
    ADVANCE_TIME(20000000); loop();
    ADVANCE_TIME(20000000); loop();
    ADVANCE_TIME(20000000); loop();
    ADVANCE_TIME(20000000); loop();
    ADVANCE_TIME(20000000); loop();
    ADVANCE_TIME(20000000); loop();
    ADVANCE_TIME(20000000); loop();
    ADVANCE_TIME(20000000); loop();
    ADVANCE_TIME(20000000); loop();
    ADVANCE_TIME(20000000); loop();
    ADVANCE_TIME(20000000); loop();
    ADVANCE_TIME(20000000); loop();
    ADVANCE_TIME(20000000); loop();
    ADVANCE_TIME(20000000); loop();
    ADVANCE_TIME(20000000); loop();
    ADVANCE_TIME(20000000); loop();
    ADVANCE_TIME(20000000); loop();
    ADVANCE_TIME(20000000); loop();
    ADVANCE_TIME(20000000); loop();
    ADVANCE_TIME(20000000); loop();
    ADVANCE_TIME(20000000); loop();
    ADVANCE_TIME(20000000); loop();
    ADVANCE_TIME(20000000); loop();
    ADVANCE_TIME(20000000); loop();
    ADVANCE_TIME(20000000); loop();
    ADVANCE_TIME(20000000); loop();
    ADVANCE_TIME(20000000); loop();
    ADVANCE_TIME(20000000); loop();
    ADVANCE_TIME(20000000); loop();
    ADVANCE_TIME(20000000); loop();
    ADVANCE_TIME(20000000); loop();
    ADVANCE_TIME(20000000); loop();
    ADVANCE_TIME(20000000); loop();
    ADVANCE_TIME(20000000); loop();
    ADVANCE_TIME(20000000); loop();
    ADVANCE_TIME(20000000); loop();
    ADVANCE_TIME(20000000); loop();
    ADVANCE_TIME(20000000); loop();
    ADVANCE_TIME(20000000); loop();
    ADVANCE_TIME(20000000); loop();
    ADVANCE_TIME(20000000); loop();
    ADVANCE_TIME(20000000); loop();
    ADVANCE_TIME(20000000); loop();
    ADVANCE_TIME(20000000); loop();
    ADVANCE_TIME(20000000); loop();
    ADVANCE_TIME(20000000); loop();
    ADVANCE_TIME(20000000); loop();
    ADVANCE_TIME(20000000); loop();
    ADVANCE_TIME(20000000); loop();
    ADVANCE_TIME(20000000); loop();
    ADVANCE_TIME(20000000); loop();
    ADVANCE_TIME(20000000); loop();
    ADVANCE_TIME(20000000); loop();
    ADVANCE_TIME(20000000); loop();
    ADVANCE_TIME(20000000); loop();
    ADVANCE_TIME(20000000); loop();
    ADVANCE_TIME(20000000); loop();
    ADVANCE_TIME(20000000); loop();
    ADVANCE_TIME(20000000); loop();
    ADVANCE_TIME(20000000); loop();
    ADVANCE_TIME(20000000); loop();
    ADVANCE_TIME(20000000); loop();
    ADVANCE_TIME(20000000); loop();
    ADVANCE_TIME(20000000); loop();
    ADVANCE_TIME(20000000); loop();
    ADVANCE_TIME(20000000); loop();
    ADVANCE_TIME(20000000); loop();
    ADVANCE_TIME(20000000); loop();
    ADVANCE_TIME(20000000); loop();
    ADVANCE_TIME(20000000); loop();
    ADVANCE_TIME(20000000); loop();
    ADVANCE_TIME(20000000); loop();
    ADVANCE_TIME(20000000); loop();
    ADVANCE_TIME(20000000); loop();
    ADVANCE_TIME(20000000); loop();
    ADVANCE_TIME(20000000); loop();
    ADVANCE_TIME(20000000); loop();
    ADVANCE_TIME(20000000); loop();
    ADVANCE_TIME(20000000); loop();
    ADVANCE_TIME(20000000); loop();
    ADVANCE_TIME(20000000); loop();
    ADVANCE_TIME(20000000); loop();
    ADVANCE_TIME(20000000); loop();
    ADVANCE_TIME(20000000); loop();
    ADVANCE_TIME(20000000); loop();
    ADVANCE_TIME(20000000); loop();
    ADVANCE_TIME(20000000); loop();
    ADVANCE_TIME(20000000); loop();
    ADVANCE_TIME(20000000); loop();
    ADVANCE_TIME(20000000); loop();
    ADVANCE_TIME(20000000); loop();
    ADVANCE_TIME(20000000); loop();
    ADVANCE_TIME(20000000); loop();
    ADVANCE_TIME(20000000); loop();
    ADVANCE_TIME(20000000); loop();
    ADVANCE_TIME(20000000); loop();
    ADVANCE_TIME(20000000); loop();
    ADVANCE_TIME(20000000); loop();
    ADVANCE_TIME(20000000); loop();
    ADVANCE_TIME(20000000); loop();
    ADVANCE_TIME(20000000); loop();
    ADVANCE_TIME(20000000); loop();
    ADVANCE_TIME(20000000); loop();
    ADVANCE_TIME(20000000); loop();
    ADVANCE_TIME(20000000); loop();
    ADVANCE_TIME(20000000); loop();
    ADVANCE_TIME(20000000); loop();
    ADVANCE_TIME(20000000); loop();
    ADVANCE_TIME(20000000); loop();
    ADVANCE_TIME(20000000); loop();
    ADVANCE_TIME(20000000); loop();
    ADVANCE_TIME(20000000); loop();
    ADVANCE_TIME(20000000); loop();
    ADVANCE_TIME(20000000); loop();
    ADVANCE_TIME(20000000); loop();
    ADVANCE_TIME(20000000); loop();
    ADVANCE_TIME(20000000); loop();
    ASSERT_EQ(loop.Phase, 3, 'Scenario termine (arret apres P1)');
    ASSERT_NEAR(loop.FreqAtCross_Hz, 20.0, 0.5, 'Approche a 20 Hz au franchissement de P1');
    ASSERT_NEAR(loop.MaxCmdAfter_Hz, 20.0, 0.5, 'Demande tenue : la consigne vers le variateur reste plafonnee a 20 Hz apres P1');
    ASSERT_GE(loop.Overshoot_M, 0.30, 'Depassement apres P1 >= 0,30 m (caracterisation)');
    ASSERT_LE(loop.Overshoot_M, 0.80, 'Depassement apres P1 <= 0,80 m (caracterisation)');
END_TEST
